   // ---------- 网络 6 ----------
   // 标题：模式传递到M区,方便使用
   // 含义：当 #SubSysMode.Mode.ManMode 为 TRUE 时置位 "ManMode_M"，否则复位（触点→线圈）
   IF #SubSysMode.Mode.ManMode THEN
       "ManMode_M" := TRUE;
   ELSE
       "ManMode_M" := FALSE;
   END_IF;
   // 含义：当 #SubSysMode.Mode.ManMode 为 TRUE 时置位 "DB1900_Communication_PC".Send.ManMode，否则复位（触点→线圈）
   IF #SubSysMode.Mode.ManMode THEN
       "DB1900_Communication_PC".Send.ManMode := TRUE;
   ELSE
       "DB1900_Communication_PC".Send.ManMode := FALSE;
   END_IF;
   // 含义：当 #SubSysMode.Mode.MastMode 为 TRUE 时置位 "MastMode_M"，否则复位（触点→线圈）
   IF #SubSysMode.Mode.MastMode THEN
       "MastMode_M" := TRUE;
   ELSE
       "MastMode_M" := FALSE;
   END_IF;
   // 含义：当 #SubSysMode.Mode.StepMode 为 TRUE 时置位 "StepMode_M"，否则复位（触点→线圈）
   IF #SubSysMode.Mode.StepMode THEN
       "StepMode_M" := TRUE;
   ELSE
       "StepMode_M" := FALSE;
   END_IF;
   // 含义：当 #SubSysMode.Mode.AutoMode 为 TRUE 时置位 "AutoMode_M"，否则复位（触点→线圈）
   IF #SubSysMode.Mode.AutoMode THEN
       "AutoMode_M" := TRUE;
   ELSE
       "AutoMode_M" := FALSE;
   END_IF;
   // 含义：当 #SubSysMode.Mode.AutoMode 为 TRUE 时置位 "DB1900_Communication_PC".Send.AutoMode，否则复位（触点→线圈）
   IF #SubSysMode.Mode.AutoMode THEN
       "DB1900_Communication_PC".Send.AutoMode := TRUE;
   ELSE
       "DB1900_Communication_PC".Send.AutoMode := FALSE;
   END_IF;
   // 含义：当 #SubSysMode.Mode.EMMode 为 TRUE 时置位 "EMMode_M"，否则复位（触点→线圈）
   IF #SubSysMode.Mode.EMMode THEN
       "EMMode_M" := TRUE;
   ELSE
       "EMMode_M" := FALSE;
   END_IF;
   // 含义：当 #SubSysMode.Mode.EMMode 为 TRUE 时置位 "DB1900_Communication_PC".Send.EmmMode，否则复位（触点→线圈）
   IF #SubSysMode.Mode.EMMode THEN
       "DB1900_Communication_PC".Send.EmmMode := TRUE;
   ELSE
       "DB1900_Communication_PC".Send.EmmMode := FALSE;
   END_IF;
   // 含义：当 #SubSysMode.Mode.StepPls 为 TRUE 时置位 "StepPls_M"，否则复位（触点→线圈）
   IF #SubSysMode.Mode.StepPls THEN
       "StepPls_M" := TRUE;
   ELSE
       "StepPls_M" := FALSE;
   END_IF;
   // 含义：当 #SubSysMode.Status.AutoModeStarted 为 TRUE 时置位 "AutoModeStarted_M"，否则复位（触点→线圈）
   IF #SubSysMode.Status.AutoModeStarted THEN
       "AutoModeStarted_M" := TRUE;
   ELSE
       "AutoModeStarted_M" := FALSE;
   END_IF;
   // 含义：当 #SubSysMode.Mode.ASMode 为 TRUE 时置位 "ASMode_M"，否则复位（触点→线圈）
   IF #SubSysMode.Mode.ASMode THEN
       "ASMode_M" := TRUE;
   ELSE
       "ASMode_M" := FALSE;
   END_IF;
   // 含义：当 #SubSysMode.Mode.ASMMode 为 TRUE 时置位 "ASMMode_M"，否则复位（触点→线圈）
   IF #SubSysMode.Mode.ASMMode THEN
       "ASMMode_M" := TRUE;
   ELSE
       "ASMMode_M" := FALSE;
   END_IF;
   // 含义：当 #SubSysMode.Mode.AllMode 为 TRUE 时置位 "AllMode_M"，否则复位（触点→线圈）
   IF #SubSysMode.Mode.AllMode THEN
       "AllMode_M" := TRUE;
   ELSE
       "AllMode_M" := FALSE;
   END_IF;
   // 含义：当 #SubSysMode.Mode.ErrRst 为 TRUE 时置位 "ErrRst_M"，否则复位（触点→线圈）
   IF #SubSysMode.Mode.ErrRst THEN
       "ErrRst_M" := TRUE;
   ELSE
       "ErrRst_M" := FALSE;
   END_IF;
   // 含义：将 #SubSysMode.Mode.ErrRst OR "DB1010_Parameter".SystemParaR.bit.ErrAutoResetOption 赋给 "ErrRst_M_Auto"
   "ErrRst_M_Auto" := #SubSysMode.Mode.ErrRst OR "DB1010_Parameter".SystemParaR.bit.ErrAutoResetOption;
   // 含义：当 "DB1010_Parameter".SystemParaR.bit.MESActive 为 TRUE 时置位 "MESConnect"，否则复位（触点→线圈）
   IF "DB1010_Parameter".SystemParaR.bit.MESActive THEN
       "MESConnect" := TRUE;
   ELSE
       "MESConnect" := FALSE;
   END_IF;

   // ---------- 网络 7 ----------
   // 标题：操作盒急停OK
   // 含义：当 NOT ("IEMOK1") 为 TRUE 时置位 "DB1148_PromptBeeper".Public.EMOK，否则复位（触点→线圈）
   IF NOT ("IEMOK1") THEN
       "DB1148_PromptBeeper".Public.EMOK := TRUE;
   ELSE
       "DB1148_PromptBeeper".Public.EMOK := FALSE;
   END_IF;
   // 含义：当 NOT ("IInsideEMOK") 为 TRUE 时置位 "DB1148_PromptBeeper".Public.InsideEMOK，否则复位（触点→线圈）
   IF NOT ("IInsideEMOK") THEN
       "DB1148_PromptBeeper".Public.InsideEMOK := TRUE;
   ELSE
       "DB1148_PromptBeeper".Public.InsideEMOK := FALSE;
   END_IF;
   // 含义：当 NOT ("IInsideEMOK1") 为 TRUE 时置位 "DB1148_PromptBeeper".Public.InsideEMOK1，否则复位（触点→线圈）
   IF NOT ("IInsideEMOK1") THEN
       "DB1148_PromptBeeper".Public.InsideEMOK1 := TRUE;
   ELSE
       "DB1148_PromptBeeper".Public.InsideEMOK1 := FALSE;
   END_IF;
   // 含义：当 NOT ("IRobotEMOK") 为 TRUE 时置位 "DB1148_PromptBeeper".Public.RobotEMOK，否则复位（触点→线圈）
   IF NOT ("IRobotEMOK") THEN
       "DB1148_PromptBeeper".Public.RobotEMOK := TRUE;
   ELSE
       "DB1148_PromptBeeper".Public.RobotEMOK := FALSE;
   END_IF;

   // ---------- 网络 8 ----------
   // 标题：调试的时候，临时关闭
   // 含义：条件 "EMMode_M" OR "DB1010_Parameter".Status.Para_ReNewEdPls OR "DB1000_StdSignal".PLS.InitialPls 成立时，将 FALSE 传送到 "Debug_True"
   IF "EMMode_M" OR "DB1010_Parameter".Status.Para_ReNewEdPls OR "DB1000_StdSignal".PLS.InitialPls THEN
       "Debug_True" := FALSE;
   END_IF;
END_FUNCTION_BLOCK

FUNCTION_BLOCK "FB1002_subSysMode"   // FB1002, SCL
{ S7_Optimized_Access := 'TRUE' }
// ============================================================
//  Block: FB1002_subSysMode
//  ============================================================
//  编号：FB1002
//  原始语言：LAD（规则翻译为 SCL）
//  含义：故障红色指示灯输出，并且存储最后的不合格状态。
   VAR_INPUT
      I_OkToStartNew : Bool;   // 可以启动新的流程
      iEMOK : Bool;   // 紧急停止OK信号
      iAirPressOK : Bool;   // 气源OK信号
      iManMode : Bool;   // 手动模式
      iAutoMode : Bool;   // 自动模式信号
      iAutoModeStart : Bool;   // 自动模式启动开关
      iBeeperQuiet : Bool;   // 蜂鸣器静音按钮
      iErrRst : Bool;   // 故障复位按钮
      iStartL : Bool;   // 左启动
      iStartR : Bool;   // 右启动
      I_ErrPresent : Bool;   // DB_ERR内有故障位存在
      I_ErrAutoReset : Bool := TRUE;   // 故障发生后自动复位。
      I_AutoRuning : Bool;   // 设备自动运行中
      I_HomeIng : Bool;   // 设备正在回原点
      I_AllStationInHomePos : Bool;   // 都在原点位置
      iHomeMode : Bool;   // 回原点按钮
      I_SP2 : Bool;   // 输入参数
   END_VAR
   VAR_OUTPUT
      oTLBlue : Bool;   // 通讯正常 塔灯-蓝
      oTLYel : Bool;   // 手动模式 塔灯-黄
      oTLGreen : Bool;   // 自动运行 塔灯-绿
      oTLRed : Bool;   // 故障报警 塔灯-红
      oTLWhite : Bool;   // 设备上电 塔灯-白
      oPanelG : Bool;   // 面板绿灯
      oPanelRed : Bool;   // 面板红灯
      oBeeper : Bool;   // 蜂鸣器
      oLightingLampClose : Bool;   // 日光灯控制
      oEMErr : Bool;   // 紧急停止故障
      oPressErr : Bool;   // 气压低故障
      oErrToBeRst : Bool;   // 发生故障，需要复位，用于屏幕提示
      oStartAutoModePrompt : Bool;   // 请启动自动模式
      oAutoModeOffPrompt : Bool;   // 自动模式已经暂停，等待循环结束！
      oEmptyMode : Bool;   // 设备进入清空模式提示信息
      oStepMode : Bool;   // 设备进入单步模式提示信息
      oModeFromTP : Bool;   // 模式来自触摸屏提示信息！
   END_VAR
   VAR
      OUT : Struct   // 静态变量
         LampTest : Bool;   // 指示灯测试
         oPanelHome : Bool;   // 面板回原点指示灯
         sp : Word;   // 静态变量
      END_STRUCT;
      Mode : Struct   // 静态变量
         ManMode : Bool;   // 手动模式
         MastMode : Bool;   // 校验模式
         StepMode : Bool;   // 单步模式
         AutoMode : Bool;   // 自动模式
         EMMode : Bool;   // 紧急停止模式
         PressLowMode : Bool;   // 气压低
         sp_1 : Bool;   // 静态变量
         sp_2 : Bool;   // 静态变量
         ASMode : Bool;   // 自动或单步模式
         ASMMode : Bool;   // 自动，单步，校验模式
         AllMode : Bool;   // 所有模式
         HomeCmd : Bool;   // 回原点命令
         ErrRst : Bool;   // 故障复位（含TPPB）
         StartPls : Bool;   // 双手启动模式使用
         StepPls : Bool;   // 双手启动模式使用
         StartLeftPls : Bool;   // 单手启动左工位
         StartRightPls : Bool;   // 单手启动右工位
         StepLeftPls : Bool;   // 单手启动左工位
         StepRightPls : Bool;   // 单手启动右工位
         ManModePls : Bool;   // 切换到手动模式脉冲
         AllModePls : Bool;   // 模式切换脉冲
         sp : DWord;   // 静态变量
      END_STRUCT;
      TPPB : Struct   // 18
         EmptyMode : Bool;   // 清空模式开始
         Bypass : Bool;   // 静态变量
         STAT6 : Bool;   // 静态变量
         STAT5 : Bool;   // 静态变量
         STAT4 : Bool;   // 静态变量
         STAT3 : Bool;   // 静态变量
         STAT2 : Bool;   // 静态变量
         STAT1 : Bool;   // 静态变量
         LampTest : Bool;   // 指示灯测试
         Home : Bool;   // 回原点
         StepMode : Bool;   // 单步按钮
         ErrRst : Bool;   // 来自触摸屏
         LampCtrol : Bool;   // ON,日光灯开
         Quiet : Bool;   // 静音，蜂鸣器
         opModeFromTP : Bool;   // 工作模式来自触摸屏选项
         sp : DWord;   // 静态变量
      END_STRUCT;
      AtTPPB : Word;   // 静态变量
      Status : Struct   // For_TP_Show
         HomePos : Bool;   // 在原点位置
         HomeIng : Bool;   // 正在原点
         AutoRunning : Bool;   // 自动运行中
         ErrPresent : Bool;   // 设备有故障
         AutoModeStarted : Bool;   // 自动模式已经启动！
      END_STRUCT;
      TPSetPageNo : Int;   // 设置当前画面号
      TPCurPageType : Int;   // 当前画面类型（工位分类）
      TPCurSubPage : Int;   // 画面子类型（手动、自动等）
      IO_FromTP : Struct   // 来自触摸屏的模拟仿真按钮输入
         spbyte : Byte;   // 来自触摸屏的模拟仿真按钮输入
         EMOK : Bool := TRUE;   // 紧急停止OK信号
         AirPressOK : Bool := TRUE;   // 气源OK信号
         ManMode : Bool;   // 手动模式
         AutoMode : Bool;   // 自动模式信号
         AutoModeStart : Bool;   // 自动模式启动开关
         ErrRst : Bool;   // 故障复位按钮
         StartLeft : Bool;   // 启动设备（左按钮）
         StartRight : Bool;   // 启动设备（右按钮）
      END_STRUCT;
      IO_Cur : Struct   // 当前实际使用的信号状态
         spbyte : Byte;   // 静态变量
         EMOK : Bool;   // 紧急停止OK信号
         AirPressOK : Bool;   // 气源OK信号
         ManMode : Bool;   // 手动模式
         AutoMode : Bool;   // 自动模式信号
         AutoModeStart : Bool;   // 自动模式启动开关
         ErrRst : Bool;   // 故障复位按钮
         StartLeft : Bool;   // 启动设备（左按钮）
         StartRight : Bool;   // 启动设备（右按钮）
      END_STRUCT;
      ModeDT : Struct   // 模式延时
         ManMode1 : Bool;   // 静态变量
         ManMode2 : Bool;   // 静态变量
         AutoMode1 : Bool;   // 静态变量
         AutoMode2 : Bool;   // 静态变量
         MastMode1 : Bool;   // 静态变量
         MastMode2 : Bool;   // 静态变量
         HomeCmd1 : Bool;   // 静态变量
         HomeCmd2 : Bool;   // 静态变量
         HomeCmd3 : Bool;   // 静态变量
         HomeCmd4 : Bool;   // 静态变量
         ErrLampOn01 : Bool;   // 静态变量
         ErrLampOn02 : Bool;   // 静态变量
      END_STRUCT;
      Aux : Struct   // 静态变量
         BeeperON_Keep : Bool;   // 静态变量
         BeeperOn : Bool;   // 静态变量
         BeeperOnPls : Bool;   // 静态变量
         ManMode : Bool;   // 用于清除触摸屏的模式选择
         ManModePls : Bool;   // 用于清除触摸屏的模式选择
         AutoMode : Bool;   // 用于清除触摸屏的模式选择
         AutoModePls : Bool;   // 用于清除触摸屏的模式选择
         ModeChangePlsHW : Bool;   // 用于记录节拍
         AutoRunningPls : Bool;   // 用于记录节拍
         OKPartPromptPls : Bool;   // 脉冲计数用
         NGPartPromptPls : Bool;   // 脉冲计数用
         ManModeOn : Bool;   // 静态变量
         AllModeOn : Bool;   // 静态变量
         AutoModeStartBtnPls : Bool;   // 静态变量
         AutoModeOnPls : Bool;   // 静态变量
         AutoModeOffCmd : Bool;   // 静态变量
         TPCurSubPage : Int;   // 静态变量
      END_STRUCT;
      Start1DT1 : IEC_TIMER;   // 静态变量
      Start1DT2 : IEC_TIMER;   // 静态变量
      Start2DT1 : IEC_TIMER;   // 静态变量
      Start2DT2 : IEC_TIMER;   // 静态变量
      xArray_SP : Array[0..91] of Byte;   // 静态变量
      lastByteAddr : Byte := 198;   // 198
      PT : Time;   // 静态变量
      ET : Time;   // 静态变量
      IN : Bool;   // 静态变量
      Q : Bool;   // 静态变量
   END_VAR
   VAR_TEMP
      T_INT : Int;   // 临时变量
   END_VAR
BEGIN

   // ---------- 网络 1 ----------
   // 标题：模拟仿真模式按钮等
   // 含义：将 (NOT (#TPPB.opModeFromTP) AND #iEMOK) OR (#TPPB.opModeFromTP AND #IO_FromTP.EMOK) 赋给 #IO_Cur.EMOK
   #IO_Cur.EMOK := (NOT (#TPPB.opModeFromTP) AND #iEMOK) OR (#TPPB.opModeFromTP AND #IO_FromTP.EMOK);
   // 含义：将 (NOT (#TPPB.opModeFromTP) AND #iAirPressOK) OR (#TPPB.opModeFromTP AND #IO_FromTP.AirPressOK) 赋给 #IO_Cur.AirPressOK
   #IO_Cur.AirPressOK := (NOT (#TPPB.opModeFromTP) AND #iAirPressOK) OR (#TPPB.opModeFromTP AND #IO_FromTP.AirPressOK);
   // 含义：将 (NOT (#TPPB.opModeFromTP) AND #iManMode) OR (#TPPB.opModeFromTP AND NOT (#IO_FromTP.AutoMode)) 赋给 #IO_Cur.ManMode
   #IO_Cur.ManMode := (NOT (#TPPB.opModeFromTP) AND #iManMode) OR (#TPPB.opModeFromTP AND NOT (#IO_FromTP.AutoMode));
   // 含义：将 (NOT (#TPPB.opModeFromTP) AND #iAutoMode) OR (#TPPB.opModeFromTP AND #IO_FromTP.AutoMode) 赋给 #IO_Cur.AutoMode
   #IO_Cur.AutoMode := (NOT (#TPPB.opModeFromTP) AND #iAutoMode) OR (#TPPB.opModeFromTP AND #IO_FromTP.AutoMode);
   // 含义：将 (NOT (#TPPB.opModeFromTP) AND #iAutoModeStart) OR (#TPPB.opModeFromTP AND #IO_FromTP.AutoModeStart) 赋给 #IO_Cur.AutoModeStart
   #IO_Cur.AutoModeStart := (NOT (#TPPB.opModeFromTP) AND #iAutoModeStart) OR (#TPPB.opModeFromTP AND #IO_FromTP.AutoModeStart);
   // 含义：将 (NOT (#TPPB.opModeFromTP) AND #iErrRst) OR (#TPPB.opModeFromTP AND #IO_FromTP.ErrRst) 赋给 #IO_Cur.ErrRst
   #IO_Cur.ErrRst := (NOT (#TPPB.opModeFromTP) AND #iErrRst) OR (#TPPB.opModeFromTP AND #IO_FromTP.ErrRst);
   // 含义：将 (NOT (#TPPB.opModeFromTP) AND #iStartL) OR (#TPPB.opModeFromTP AND #IO_FromTP.StartLeft) 赋给 #IO_Cur.StartLeft
   #IO_Cur.StartLeft := (NOT (#TPPB.opModeFromTP) AND #iStartL) OR (#TPPB.opModeFromTP AND #IO_FromTP.StartLeft);
   // 含义：将 (NOT (#TPPB.opModeFromTP) AND #iStartR) OR (#TPPB.opModeFromTP AND #IO_FromTP.StartRight) 赋给 #IO_Cur.StartRight
   #IO_Cur.StartRight := (NOT (#TPPB.opModeFromTP) AND #iStartR) OR (#TPPB.opModeFromTP AND #IO_FromTP.StartRight);
   // 含义：条件 (#iManMode OR #iAutoMode) AND NOT (#Aux.ModeChangePlsHW) 成立时，将 FALSE 传送到 #TPPB.opModeFromTP
   IF (#iManMode OR #iAutoMode) AND NOT (#Aux.ModeChangePlsHW) THEN
       #TPPB.opModeFromTP := FALSE;
   END_IF;
   // 含义：将 #iManMode OR #iAutoMode 赋给 #Aux.ModeChangePlsHW
   #Aux.ModeChangePlsHW := #iManMode OR #iAutoMode;
   // 含义：当 #TPPB.opModeFromTP 为 TRUE 时置位 #oModeFromTP，否则复位（触点→线圈）
   IF #TPPB.opModeFromTP THEN
       #oModeFromTP := TRUE;
   ELSE
       #oModeFromTP := FALSE;
   END_IF;
   // 含义：条件 #TPPB.opModeFromTP AND #iErrRst 成立时，将 FALSE 传送到 #TPPB.opModeFromTP
   IF #TPPB.opModeFromTP AND #iErrRst THEN
       #TPPB.opModeFromTP := FALSE;
   END_IF;

   // ---------- 网络 2 ----------
   // 标题：在原点位置
   // 含义：当 #I_AllStationInHomePos 为 TRUE 时置位 #Status.HomePos，否则复位（触点→线圈）
   IF #I_AllStationInHomePos THEN
       #Status.HomePos := TRUE;
   ELSE
       #Status.HomePos := FALSE;
   END_IF;
   // 含义：当 #I_HomeIng 为 TRUE 时置位 #Status.HomeIng，否则复位（触点→线圈）
   IF #I_HomeIng THEN
       #Status.HomeIng := TRUE;
   ELSE
       #Status.HomeIng := FALSE;
   END_IF;
   // 含义：当 #I_AutoRuning 为 TRUE 时置位 #Status.AutoRunning，否则复位（触点→线圈）
   IF #I_AutoRuning THEN
       #Status.AutoRunning := TRUE;
   ELSE
       #Status.AutoRunning := FALSE;
   END_IF;

   // ---------- 网络 3 ----------
   // 标题：#OUT.ErrLamp
   // 含义：当 #I_ErrPresent 为 TRUE 时置位 #Status.ErrPresent，否则复位（触点→线圈）
   IF #I_ErrPresent THEN
       #Status.ErrPresent := TRUE;
   ELSE
       #Status.ErrPresent := FALSE;
   END_IF;

   // ---------- 网络 4 ----------
   // 标题：#oTLRed
   // 注释：故障红色指示灯输出，并且存储最后的不合格状态。
   // 含义：将 #Status.ErrPresent AND #ModeDT.ErrLampOn02 赋给 #oTLRed
   #oTLRed := #Status.ErrPresent AND #ModeDT.ErrLampOn02;
   // 含义：将 ((#Status.ErrPresent AND "DB1000_StdSignal".PLS.PS05) AND #ModeDT.ErrLampOn01) OR (#Status.ErrPresent AND #ModeDT.ErrLampOn02) 赋给 #ModeDT.ErrLampOn02
   #ModeDT.ErrLampOn02 := ((#Status.ErrPresent AND "DB1000_StdSignal".PLS.PS05) AND #ModeDT.ErrLampOn01) OR (#Status.ErrPresent AND #ModeDT.ErrLampOn02);
   // 含义：将 (#Status.ErrPresent AND "DB1000_StdSignal".PLS.PS01) OR (#Status.ErrPresent AND #ModeDT.ErrLampOn01) 赋给 #ModeDT.ErrLampOn01
   #ModeDT.ErrLampOn01 := (#Status.ErrPresent AND "DB1000_StdSignal".PLS.PS01) OR (#Status.ErrPresent AND #ModeDT.ErrLampOn01);

   // ---------- 网络 5 ----------
   // 标题：#oTLYel,   #oTLGreen
   // 含义：当 #Mode.ManMode 为 TRUE 时置位 #oTLYel，否则复位（触点→线圈）
   IF #Mode.ManMode THEN
       #oTLYel := TRUE;
   ELSE
       #oTLYel := FALSE;
   END_IF;
   // 含义：将 #Mode.ASMMode AND NOT (#oTLRed) 赋给 #oTLGreen
   #oTLGreen := #Mode.ASMMode AND NOT (#oTLRed);

   // ---------- 网络 6 ----------
   // 标题：#oTLBlue
   // 含义：将 "DB720_KuKa_MainCtrl".ChangeTool.StepStart AND "DB1000_StdSignal".RectWave.Wave05 赋给 #oTLBlue
   #oTLBlue := "DB720_KuKa_MainCtrl".ChangeTool.StepStart AND "DB1000_StdSignal".RectWave.Wave05;
   // 含义：当 NOT (#Mode.EMMode) 为 TRUE 时置位 #oTLWhite，否则复位（触点→线圈）
   IF NOT (#Mode.EMMode) THEN
       #oTLWhite := TRUE;
   ELSE
       #oTLWhite := FALSE;
   END_IF;

   // ---------- 网络 7 ----------
   // 标题：#oPanelG
   // 含义：将 ((((#Status.HomeIng AND "DB1000_StdSignal".RectWave.Wave02) AND NOT (TRUE)) OR (((((#Mode.AutoMode AND NOT (#I_HomeIng)) AND NOT (#Status.AutoRunning)) AND NOT (#Status.AutoModeStarted)) AND #Status.HomePos) AND "DB1000_StdSignal".RectWave.Wave05) OR #Status.AutoModeStarted OR ("AutoMode_M" AND "DB1900_Communication_PC".Send.DrillRunning)) AND NOT (#Aux.AutoModeOffCmd)) OR (#Aux.AutoModeOffCmd AND "DB1000_StdSignal".PLS.PS02) 赋给 #oPanelG
   #oPanelG := ((((#Status.HomeIng AND "DB1000_StdSignal".RectWave.Wave02) AND NOT (TRUE)) OR (((((#Mode.AutoMode AND NOT (#I_HomeIng)) AND NOT (#Status.AutoRunning)) AND NOT (#Status.AutoModeStarted)) AND #Status.HomePos) AND "DB1000_StdSignal".RectWave.Wave05) OR #Status.AutoModeStarted OR ("AutoMode_M" AND "DB1900_Communication_PC".Send.DrillRunning)) AND NOT (#Aux.AutoModeOffCmd)) OR (#Aux.AutoModeOffCmd AND "DB1000_StdSignal".PLS.PS02);

   // ---------- 网络 8 ----------
   // 标题：#oPanelRed
   // 注释：故障红色指示灯输出，并且存储最后的不合格状态。
   // 含义：将 #oTLRed OR (#I_HomeIng AND "DB1000_StdSignal".RectWave.Wave02) 赋给 #oPanelRed
   #oPanelRed := #oTLRed OR (#I_HomeIng AND "DB1000_StdSignal".RectWave.Wave02);

   // ---------- 网络 9 ----------
   // 标题：#oBeeper
   // 含义：将 #oTLRed AND NOT (#Aux.BeeperOn) 赋给 #Aux.BeeperOnPls
   #Aux.BeeperOnPls := #oTLRed AND NOT (#Aux.BeeperOn);
   // 含义：当 #oTLRed 为 TRUE 时置位 #Aux.BeeperOn，否则复位（触点→线圈）
   IF #oTLRed THEN
       #Aux.BeeperOn := TRUE;
   ELSE
       #Aux.BeeperOn := FALSE;
   END_IF;
   // 含义：将 (((#oTLRed AND #Aux.BeeperOnPls) OR (#oTLRed AND #Aux.BeeperON_Keep)) AND NOT (#Mode.ErrRst)) AND NOT (#iBeeperQuiet) 赋给 #Aux.BeeperON_Keep
   #Aux.BeeperON_Keep := (((#oTLRed AND #Aux.BeeperOnPls) OR (#oTLRed AND #Aux.BeeperON_Keep)) AND NOT (#Mode.ErrRst)) AND NOT (#iBeeperQuiet);
   // 含义：将 (((#oTLRed AND #Aux.BeeperOnPls) OR (#oTLRed AND #Aux.BeeperON_Keep)) AND "DB1000_StdSignal".RectWave.Beeper) AND NOT (#TPPB.Quiet) 赋给 #oBeeper
   #oBeeper := (((#oTLRed AND #Aux.BeeperOnPls) OR (#oTLRed AND #Aux.BeeperON_Keep)) AND "DB1000_StdSignal".RectWave.Beeper) AND NOT (#TPPB.Quiet);

   // ---------- 网络 10 ----------
   // 标题：#oPanelHome
   // 含义：将 (#Status.HomeIng AND "DB1000_StdSignal".RectWave.Wave02) OR #I_AllStationInHomePos 赋给 #OUT.oPanelHome
   #OUT.oPanelHome := (#Status.HomeIng AND "DB1000_StdSignal".RectWave.Wave02) OR #I_AllStationInHomePos;

   // ---------- 网络 11 ----------
   // 标题：#oErrToBeRst
   // 含义：将 (((#oTLRed OR #oErrToBeRst) AND NOT (#Mode.ErrRst)) AND NOT (#I_ErrAutoReset)) AND #Mode.AllMode 赋给 #oErrToBeRst
   #oErrToBeRst := (((#oTLRed OR #oErrToBeRst) AND NOT (#Mode.ErrRst)) AND NOT (#I_ErrAutoReset)) AND #Mode.AllMode;

   // ---------- 网络 12 ----------
   // 标题：#oEMErr,   #oPressErr
   // 含义：当 NOT (#IO_Cur.EMOK) 为 TRUE 时置位 #oEMErr，否则复位（触点→线圈）
   IF NOT (#IO_Cur.EMOK) THEN
       #oEMErr := TRUE;
   ELSE
       #oEMErr := FALSE;
   END_IF;
   // 含义：条件 #IO_Cur.EMOK AND NOT (#IO_Cur.AirPressOK) 成立时，将 TRUE 传送到 #oPressErr
   IF #IO_Cur.EMOK AND NOT (#IO_Cur.AirPressOK) THEN
       #oPressErr := TRUE;
   END_IF;
   // 含义：条件 #Mode.ErrRst AND #IO_Cur.AirPressOK 成立时，将 FALSE 传送到 #oPressErr
   IF #Mode.ErrRst AND #IO_Cur.AirPressOK THEN
       #oPressErr := FALSE;
   END_IF;

   // ---------- 网络 13 ----------
   // 标题：Mode ChangePls;
   // 含义：将 #IO_Cur.ManMode AND NOT (#Aux.ManMode) 赋给 #Aux.ManModePls
   #Aux.ManModePls := #IO_Cur.ManMode AND NOT (#Aux.ManMode);
   // 含义：当 #IO_Cur.ManMode 为 TRUE 时置位 #Aux.ManMode，否则复位（触点→线圈）
   IF #IO_Cur.ManMode THEN
       #Aux.ManMode := TRUE;
   ELSE
       #Aux.ManMode := FALSE;
   END_IF;
   // 含义：将 #IO_Cur.AutoMode AND NOT (#Aux.AutoMode) 赋给 #Aux.AutoModePls
   #Aux.AutoModePls := #IO_Cur.AutoMode AND NOT (#Aux.AutoMode);
   // 含义：当 #IO_Cur.AutoMode 为 TRUE 时置位 #Aux.AutoMode，否则复位（触点→线圈）
   IF #IO_Cur.AutoMode THEN
       #Aux.AutoMode := TRUE;
   ELSE
       #Aux.AutoMode := FALSE;
   END_IF;

   // ---------- 网络 14 ----------
   // 标题：模式延时处理。
   // 含义：将 (((((("DB1000_StdSignal".PowerOn AND NOT (#oEMErr)) AND NOT (#oPressErr)) AND #IO_Cur.ManMode) AND NOT (#IO_Cur.AutoMode)) AND "DB1000_StdSignal".PLS.PS01) AND #ModeDT.ManMode1) OR ((((("DB1000_StdSignal".PowerOn AND NOT (#oEMErr)) AND NOT (#oPressErr)) AND #IO_Cur.ManMode) AND NOT (#IO_Cur.AutoMode)) AND #ModeDT.ManMode2) 赋给 #ModeDT.ManMode2
   #ModeDT.ManMode2 := (((((("DB1000_StdSignal".PowerOn AND NOT (#oEMErr)) AND NOT (#oPressErr)) AND #IO_Cur.ManMode) AND NOT (#IO_Cur.AutoMode)) AND "DB1000_StdSignal".PLS.PS01) AND #ModeDT.ManMode1) OR ((((("DB1000_StdSignal".PowerOn AND NOT (#oEMErr)) AND NOT (#oPressErr)) AND #IO_Cur.ManMode) AND NOT (#IO_Cur.AutoMode)) AND #ModeDT.ManMode2);
   // 含义：将 ((((("DB1000_StdSignal".PowerOn AND NOT (#oEMErr)) AND NOT (#oPressErr)) AND #IO_Cur.ManMode) AND NOT (#IO_Cur.AutoMode)) AND "DB1000_StdSignal".PLS.PS01) OR ((((("DB1000_StdSignal".PowerOn AND NOT (#oEMErr)) AND NOT (#oPressErr)) AND #IO_Cur.ManMode) AND NOT (#IO_Cur.AutoMode)) AND #ModeDT.ManMode1) 赋给 #ModeDT.ManMode1
   #ModeDT.ManMode1 := ((((("DB1000_StdSignal".PowerOn AND NOT (#oEMErr)) AND NOT (#oPressErr)) AND #IO_Cur.ManMode) AND NOT (#IO_Cur.AutoMode)) AND "DB1000_StdSignal".PLS.PS01) OR ((((("DB1000_StdSignal".PowerOn AND NOT (#oEMErr)) AND NOT (#oPressErr)) AND #IO_Cur.ManMode) AND NOT (#IO_Cur.AutoMode)) AND #ModeDT.ManMode1);
   // 含义：将 (((((("DB1000_StdSignal".PowerOn AND NOT (#oEMErr)) AND NOT (#oPressErr)) AND NOT (#IO_Cur.ManMode)) AND #IO_Cur.AutoMode) AND "DB1000_StdSignal".PLS.PS01) AND #ModeDT.AutoMode1) OR ((((("DB1000_StdSignal".PowerOn AND NOT (#oEMErr)) AND NOT (#oPressErr)) AND NOT (#IO_Cur.ManMode)) AND #IO_Cur.AutoMode) AND #ModeDT.AutoMode2) 赋给 #ModeDT.AutoMode2
   #ModeDT.AutoMode2 := (((((("DB1000_StdSignal".PowerOn AND NOT (#oEMErr)) AND NOT (#oPressErr)) AND NOT (#IO_Cur.ManMode)) AND #IO_Cur.AutoMode) AND "DB1000_StdSignal".PLS.PS01) AND #ModeDT.AutoMode1) OR ((((("DB1000_StdSignal".PowerOn AND NOT (#oEMErr)) AND NOT (#oPressErr)) AND NOT (#IO_Cur.ManMode)) AND #IO_Cur.AutoMode) AND #ModeDT.AutoMode2);
   // 含义：将 ((((("DB1000_StdSignal".PowerOn AND NOT (#oEMErr)) AND NOT (#oPressErr)) AND NOT (#IO_Cur.ManMode)) AND #IO_Cur.AutoMode) AND "DB1000_StdSignal".PLS.PS01) OR ((((("DB1000_StdSignal".PowerOn AND NOT (#oEMErr)) AND NOT (#oPressErr)) AND NOT (#IO_Cur.ManMode)) AND #IO_Cur.AutoMode) AND #ModeDT.AutoMode1) 赋给 #ModeDT.AutoMode1
   #ModeDT.AutoMode1 := ((((("DB1000_StdSignal".PowerOn AND NOT (#oEMErr)) AND NOT (#oPressErr)) AND NOT (#IO_Cur.ManMode)) AND #IO_Cur.AutoMode) AND "DB1000_StdSignal".PLS.PS01) OR ((((("DB1000_StdSignal".PowerOn AND NOT (#oEMErr)) AND NOT (#oPressErr)) AND NOT (#IO_Cur.ManMode)) AND #IO_Cur.AutoMode) AND #ModeDT.AutoMode1);
   // 含义：将 (((((("DB1000_StdSignal".PowerOn AND NOT (#oEMErr)) AND NOT (#oPressErr)) AND NOT (#IO_Cur.ManMode)) AND NOT (#IO_Cur.AutoMode)) AND "DB1000_StdSignal".PLS.PS01) AND #ModeDT.MastMode1) OR ((((("DB1000_StdSignal".PowerOn AND NOT (#oEMErr)) AND NOT (#oPressErr)) AND NOT (#IO_Cur.ManMode)) AND NOT (#IO_Cur.AutoMode)) AND #ModeDT.MastMode2) 赋给 #ModeDT.MastMode2
   #ModeDT.MastMode2 := (((((("DB1000_StdSignal".PowerOn AND NOT (#oEMErr)) AND NOT (#oPressErr)) AND NOT (#IO_Cur.ManMode)) AND NOT (#IO_Cur.AutoMode)) AND "DB1000_StdSignal".PLS.PS01) AND #ModeDT.MastMode1) OR ((((("DB1000_StdSignal".PowerOn AND NOT (#oEMErr)) AND NOT (#oPressErr)) AND NOT (#IO_Cur.ManMode)) AND NOT (#IO_Cur.AutoMode)) AND #ModeDT.MastMode2);
   // 含义：将 ((((("DB1000_StdSignal".PowerOn AND NOT (#oEMErr)) AND NOT (#oPressErr)) AND NOT (#IO_Cur.ManMode)) AND NOT (#IO_Cur.AutoMode)) AND "DB1000_StdSignal".PLS.PS01) OR ((((("DB1000_StdSignal".PowerOn AND NOT (#oEMErr)) AND NOT (#oPressErr)) AND NOT (#IO_Cur.ManMode)) AND NOT (#IO_Cur.AutoMode)) AND #ModeDT.MastMode1) 赋给 #ModeDT.MastMode1
   #ModeDT.MastMode1 := ((((("DB1000_StdSignal".PowerOn AND NOT (#oEMErr)) AND NOT (#oPressErr)) AND NOT (#IO_Cur.ManMode)) AND NOT (#IO_Cur.AutoMode)) AND "DB1000_StdSignal".PLS.PS01) OR ((((("DB1000_StdSignal".PowerOn AND NOT (#oEMErr)) AND NOT (#oPressErr)) AND NOT (#IO_Cur.ManMode)) AND NOT (#IO_Cur.AutoMode)) AND #ModeDT.MastMode1);
   // 含义：将 (((((("DB1000_StdSignal".PowerOn AND NOT (#oEMErr)) AND NOT (#oPressErr)) AND #Mode.ErrRst) OR ((("DB1000_StdSignal".PowerOn AND NOT (#oEMErr)) AND NOT (#oPressErr)) AND #iHomeMode)) AND "DB1000_StdSignal".PLS.PS05) AND #ModeDT.HomeCmd3) OR ((((("DB1000_StdSignal".PowerOn AND NOT (#oEMErr)) AND NOT (#oPressErr)) AND #Mode.ErrRst) OR ((("DB1000_StdSignal".PowerOn AND NOT (#oEMErr)) AND NOT (#oPressErr)) AND #iHomeMode)) AND #ModeDT.HomeCmd4) 赋给 #ModeDT.HomeCmd4
   #ModeDT.HomeCmd4 := (((((("DB1000_StdSignal".PowerOn AND NOT (#oEMErr)) AND NOT (#oPressErr)) AND #Mode.ErrRst) OR ((("DB1000_StdSignal".PowerOn AND NOT (#oEMErr)) AND NOT (#oPressErr)) AND #iHomeMode)) AND "DB1000_StdSignal".PLS.PS05) AND #ModeDT.HomeCmd3) OR ((((("DB1000_StdSignal".PowerOn AND NOT (#oEMErr)) AND NOT (#oPressErr)) AND #Mode.ErrRst) OR ((("DB1000_StdSignal".PowerOn AND NOT (#oEMErr)) AND NOT (#oPressErr)) AND #iHomeMode)) AND #ModeDT.HomeCmd4);
   // 含义：将 (((((("DB1000_StdSignal".PowerOn AND NOT (#oEMErr)) AND NOT (#oPressErr)) AND #Mode.ErrRst) OR ((("DB1000_StdSignal".PowerOn AND NOT (#oEMErr)) AND NOT (#oPressErr)) AND #iHomeMode)) AND "DB1000_StdSignal".PLS.PS05) AND #ModeDT.HomeCmd2) OR ((((("DB1000_StdSignal".PowerOn AND NOT (#oEMErr)) AND NOT (#oPressErr)) AND #Mode.ErrRst) OR ((("DB1000_StdSignal".PowerOn AND NOT (#oEMErr)) AND NOT (#oPressErr)) AND #iHomeMode)) AND #ModeDT.HomeCmd3) 赋给 #ModeDT.HomeCmd3
   #ModeDT.HomeCmd3 := (((((("DB1000_StdSignal".PowerOn AND NOT (#oEMErr)) AND NOT (#oPressErr)) AND #Mode.ErrRst) OR ((("DB1000_StdSignal".PowerOn AND NOT (#oEMErr)) AND NOT (#oPressErr)) AND #iHomeMode)) AND "DB1000_StdSignal".PLS.PS05) AND #ModeDT.HomeCmd2) OR ((((("DB1000_StdSignal".PowerOn AND NOT (#oEMErr)) AND NOT (#oPressErr)) AND #Mode.ErrRst) OR ((("DB1000_StdSignal".PowerOn AND NOT (#oEMErr)) AND NOT (#oPressErr)) AND #iHomeMode)) AND #ModeDT.HomeCmd3);
   // 含义：将 (((((("DB1000_StdSignal".PowerOn AND NOT (#oEMErr)) AND NOT (#oPressErr)) AND #Mode.ErrRst) OR ((("DB1000_StdSignal".PowerOn AND NOT (#oEMErr)) AND NOT (#oPressErr)) AND #iHomeMode)) AND "DB1000_StdSignal".PLS.PS10) AND #ModeDT.HomeCmd1) OR ((((("DB1000_StdSignal".PowerOn AND NOT (#oEMErr)) AND NOT (#oPressErr)) AND #Mode.ErrRst) OR ((("DB1000_StdSignal".PowerOn AND NOT (#oEMErr)) AND NOT (#oPressErr)) AND #iHomeMode)) AND #ModeDT.HomeCmd2) 赋给 #ModeDT.HomeCmd2
   #ModeDT.HomeCmd2 := (((((("DB1000_StdSignal".PowerOn AND NOT (#oEMErr)) AND NOT (#oPressErr)) AND #Mode.ErrRst) OR ((("DB1000_StdSignal".PowerOn AND NOT (#oEMErr)) AND NOT (#oPressErr)) AND #iHomeMode)) AND "DB1000_StdSignal".PLS.PS10) AND #ModeDT.HomeCmd1) OR ((((("DB1000_StdSignal".PowerOn AND NOT (#oEMErr)) AND NOT (#oPressErr)) AND #Mode.ErrRst) OR ((("DB1000_StdSignal".PowerOn AND NOT (#oEMErr)) AND NOT (#oPressErr)) AND #iHomeMode)) AND #ModeDT.HomeCmd2);
   // 含义：将 ((((("DB1000_StdSignal".PowerOn AND NOT (#oEMErr)) AND NOT (#oPressErr)) AND #Mode.ErrRst) OR ((("DB1000_StdSignal".PowerOn AND NOT (#oEMErr)) AND NOT (#oPressErr)) AND #iHomeMode)) AND "DB1000_StdSignal".PLS.PS10) OR ((((("DB1000_StdSignal".PowerOn AND NOT (#oEMErr)) AND NOT (#oPressErr)) AND #Mode.ErrRst) OR ((("DB1000_StdSignal".PowerOn AND NOT (#oEMErr)) AND NOT (#oPressErr)) AND #iHomeMode)) AND #ModeDT.HomeCmd1) 赋给 #ModeDT.HomeCmd1
   #ModeDT.HomeCmd1 := ((((("DB1000_StdSignal".PowerOn AND NOT (#oEMErr)) AND NOT (#oPressErr)) AND #Mode.ErrRst) OR ((("DB1000_StdSignal".PowerOn AND NOT (#oEMErr)) AND NOT (#oPressErr)) AND #iHomeMode)) AND "DB1000_StdSignal".PLS.PS10) OR ((((("DB1000_StdSignal".PowerOn AND NOT (#oEMErr)) AND NOT (#oPressErr)) AND #Mode.ErrRst) OR ((("DB1000_StdSignal".PowerOn AND NOT (#oEMErr)) AND NOT (#oPressErr)) AND #iHomeMode)) AND #ModeDT.HomeCmd1);

   // ---------- 网络 15 ----------
   // 标题：AutoMode Push On
   // 含义：将 (((#Mode.ASMode AND #IO_Cur.AutoModeStart) AND NOT (#Aux.AutoModeStartBtnPls)) AND NOT (#Status.AutoModeStarted)) OR (((#Mode.ASMode AND #IO_Cur.AutoModeStart) AND NOT (#Aux.AutoModeStartBtnPls)) AND #Aux.AutoModeOffCmd) 赋给 #Aux.AutoModeOnPls
   #Aux.AutoModeOnPls := (((#Mode.ASMode AND #IO_Cur.AutoModeStart) AND NOT (#Aux.AutoModeStartBtnPls)) AND NOT (#Status.AutoModeStarted)) OR (((#Mode.ASMode AND #IO_Cur.AutoModeStart) AND NOT (#Aux.AutoModeStartBtnPls)) AND #Aux.AutoModeOffCmd);
   // 含义：条件 (((#Mode.ASMode AND #IO_Cur.AutoModeStart) AND NOT (#Aux.AutoModeStartBtnPls)) AND NOT (#Status.AutoModeStarted)) OR (((#Mode.ASMode AND #IO_Cur.AutoModeStart) AND NOT (#Aux.AutoModeStartBtnPls)) AND #Aux.AutoModeOffCmd) 成立时，将 FALSE 传送到 #Aux.AutoModeOffCmd
   IF (((#Mode.ASMode AND #IO_Cur.AutoModeStart) AND NOT (#Aux.AutoModeStartBtnPls)) AND NOT (#Status.AutoModeStarted)) OR (((#Mode.ASMode AND #IO_Cur.AutoModeStart) AND NOT (#Aux.AutoModeStartBtnPls)) AND #Aux.AutoModeOffCmd) THEN
       #Aux.AutoModeOffCmd := FALSE;
   END_IF;
   // 含义：条件 (((#Mode.ASMode AND #IO_Cur.AutoModeStart) AND NOT (#Aux.AutoModeStartBtnPls)) AND NOT (#Status.AutoModeStarted)) OR (((#Mode.ASMode AND #IO_Cur.AutoModeStart) AND NOT (#Aux.AutoModeStartBtnPls)) AND #Aux.AutoModeOffCmd) 成立时，将 FALSE 传送到 #TPPB.StepMode
   IF (((#Mode.ASMode AND #IO_Cur.AutoModeStart) AND NOT (#Aux.AutoModeStartBtnPls)) AND NOT (#Status.AutoModeStarted)) OR (((#Mode.ASMode AND #IO_Cur.AutoModeStart) AND NOT (#Aux.AutoModeStartBtnPls)) AND #Aux.AutoModeOffCmd) THEN
       #TPPB.StepMode := FALSE;
   END_IF;
   // 含义：条件 (((#Mode.ASMode AND #IO_Cur.AutoModeStart) AND NOT (#Aux.AutoModeStartBtnPls)) AND NOT (#Aux.AutoModeOnPls)) AND #Status.AutoModeStarted 成立时，将 TRUE 传送到 #Aux.AutoModeOffCmd
   IF (((#Mode.ASMode AND #IO_Cur.AutoModeStart) AND NOT (#Aux.AutoModeStartBtnPls)) AND NOT (#Aux.AutoModeOnPls)) AND #Status.AutoModeStarted THEN
       #Aux.AutoModeOffCmd := TRUE;
   END_IF;
   // 含义：将 #Mode.ASMode AND #IO_Cur.AutoModeStart 赋给 #Aux.AutoModeStartBtnPls
   #Aux.AutoModeStartBtnPls := #Mode.ASMode AND #IO_Cur.AutoModeStart;
   // 含义：将 #Mode.ASMode AND #Aux.AutoModeOffCmd 赋给 #oAutoModeOffPrompt
   #oAutoModeOffPrompt := #Mode.ASMode AND #Aux.AutoModeOffCmd;
   // 含义：条件 NOT (#Status.AutoModeStarted) AND NOT (#Status.AutoRunning) 成立时，将 FALSE 传送到 #Aux.AutoModeOffCmd
   IF NOT (#Status.AutoModeStarted) AND NOT (#Status.AutoRunning) THEN
       #Aux.AutoModeOffCmd := FALSE;
   END_IF;

   // ---------- 网络 16 ----------
   // 标题：自动模式已经启动！
   // 含义：将 (((((((#Mode.AutoMode AND #Aux.AutoModeOnPls) AND #Status.HomePos) AND #I_OkToStartNew) AND NOT (#I_AutoRuning)) AND NOT (#I_HomeIng)) OR (#Mode.AutoMode AND #Status.AutoModeStarted)) AND NOT (#TPPB.StepMode)) AND NOT (#Aux.AutoModeOffCmd) 赋给 #Status.AutoModeStarted
   #Status.AutoModeStarted := (((((((#Mode.AutoMode AND #Aux.AutoModeOnPls) AND #Status.HomePos) AND #I_OkToStartNew) AND NOT (#I_AutoRuning)) AND NOT (#I_HomeIng)) OR (#Mode.AutoMode AND #Status.AutoModeStarted)) AND NOT (#TPPB.StepMode)) AND NOT (#Aux.AutoModeOffCmd);
   // 含义：将 (#Mode.AutoMode AND NOT (#Status.AutoModeStarted)) AND NOT (#Status.AutoRunning) 赋给 #oStartAutoModePrompt
   #oStartAutoModePrompt := (#Mode.AutoMode AND NOT (#Status.AutoModeStarted)) AND NOT (#Status.AutoRunning);

   // ---------- 网络 17 ----------
   // 标题：5种模式，用于触摸屏显示
   // 含义：当 #ModeDT.ManMode2 为 TRUE 时置位 #Mode.ManMode，否则复位（触点→线圈）
   IF #ModeDT.ManMode2 THEN
       #Mode.ManMode := TRUE;
   ELSE
       #Mode.ManMode := FALSE;
   END_IF;
   // 含义：将 #ModeDT.AutoMode2 AND NOT (#TPPB.StepMode) 赋给 #Mode.AutoMode
   #Mode.AutoMode := #ModeDT.AutoMode2 AND NOT (#TPPB.StepMode);
   // 含义：将 #ModeDT.AutoMode2 AND #TPPB.StepMode 赋给 #Mode.StepMode
   #Mode.StepMode := #ModeDT.AutoMode2 AND #TPPB.StepMode;
   // 含义：当 #ModeDT.MastMode2 为 TRUE 时置位 #Mode.MastMode，否则复位（触点→线圈）
   IF #ModeDT.MastMode2 THEN
       #Mode.MastMode := TRUE;
   ELSE
       #Mode.MastMode := FALSE;
   END_IF;
   // 含义：当 #oEMErr 为 TRUE 时置位 #Mode.EMMode，否则复位（触点→线圈）
   IF #oEMErr THEN
       #Mode.EMMode := TRUE;
   ELSE
       #Mode.EMMode := FALSE;
   END_IF;
   // 含义：将 NOT (#Mode.EMMode) AND #oPressErr 赋给 #Mode.PressLowMode
   #Mode.PressLowMode := NOT (#Mode.EMMode) AND #oPressErr;

   // ---------- 网络 18 ----------
   // 标题：模式整合，用于程序中，与触摸屏无关
   // 含义：将 #Mode.AutoMode OR #Mode.StepMode 赋给 #Mode.ASMode
   #Mode.ASMode := #Mode.AutoMode OR #Mode.StepMode;
   // 含义：将 #Mode.ASMode OR #Mode.MastMode 赋给 #Mode.ASMMode
   #Mode.ASMMode := #Mode.ASMode OR #Mode.MastMode;
   // 含义：将 #Mode.ManMode OR #Mode.ASMMode 赋给 #Mode.AllMode
   #Mode.AllMode := #Mode.ManMode OR #Mode.ASMMode;
   // 含义：将 #ModeDT.HomeCmd2 OR #TPPB.Home 赋给 #Mode.HomeCmd
   #Mode.HomeCmd := #ModeDT.HomeCmd2 OR #TPPB.Home;
   // 含义：将 #IO_Cur.ErrRst OR #TPPB.ErrRst 赋给 #Mode.ErrRst
   #Mode.ErrRst := #IO_Cur.ErrRst OR #TPPB.ErrRst;

   // ---------- 网络 19 ----------
   // 标题：切换到手动模式脉冲
   // 含义：将 #Mode.ManMode AND NOT (#Aux.ManModeOn) 赋给 #Mode.ManModePls
   #Mode.ManModePls := #Mode.ManMode AND NOT (#Aux.ManModeOn);
   // 含义：当 #Mode.ManMode 为 TRUE 时置位 #Aux.ManModeOn，否则复位（触点→线圈）
   IF #Mode.ManMode THEN
       #Aux.ManModeOn := TRUE;
   ELSE
       #Aux.ManModeOn := FALSE;
   END_IF;
   // 含义：将 #Mode.AllMode AND NOT (#Aux.AllModeOn) 赋给 #Mode.AllModePls
   #Mode.AllModePls := #Mode.AllMode AND NOT (#Aux.AllModeOn);
   // 含义：当 #Mode.AllMode 为 TRUE 时置位 #Aux.AllModeOn，否则复位（触点→线圈）
   IF #Mode.AllMode THEN
       #Aux.AllModeOn := TRUE;
   ELSE
       #Aux.AllModeOn := FALSE;
   END_IF;

   // ---------- 网络 20 ----------
   // 标题：TPPB 清除；
   // 含义：条件 NOT (#Mode.AllMode) 成立时，将 FALSE 传送到 #TPPB.Home
   IF NOT (#Mode.AllMode) THEN
       #TPPB.Home := FALSE;
   END_IF;
   // 含义：条件 NOT (#Mode.AllMode) 成立时，将 FALSE 传送到 #TPPB.ErrRst
   IF NOT (#Mode.AllMode) THEN
       #TPPB.ErrRst := FALSE;
   END_IF;
   // 含义：条件 NOT (#Mode.AllMode) 成立时，将 FALSE 传送到 #TPPB.StepMode
   IF NOT (#Mode.AllMode) THEN
       #TPPB.StepMode := FALSE;
   END_IF;

   // ---------- 网络 21 ----------
   // 标题：启动延时
   // 注释：启动信号，考虑双工位情况，如果单工位，可以只用其中之一的启动，如果是双手启动
   // ，则都用上，万能！！！
   // 含义：调用计数器实例 #Start1DT1.TON（上升沿计数，当前值写入 CV）
   #Start1DT1.TON(IN := #IO_Cur.StartLeft,
                  PT := t#30ms);
   // 含义：调用计数器实例 #Start1DT2.TON（上升沿计数，当前值写入 CV）
   #Start1DT2.TON(IN := #IO_Cur.StartLeft,
                  PT := t#130ms);
   // 含义：调用计数器实例 #Start2DT1.TON（上升沿计数，当前值写入 CV）
   #Start2DT1.TON(IN := #IO_Cur.StartRight,
                  PT := t#30ms);
   // 含义：调用计数器实例 #Start2DT2.TON（上升沿计数，当前值写入 CV）
   #Start2DT2.TON(IN := #IO_Cur.StartRight,
                  PT := t#130ms);
   // 含义：将 #Start1DT1.Q AND NOT (#Start1DT2.Q) 赋给 #Mode.StartLeftPls
   #Mode.StartLeftPls := #Start1DT1.Q AND NOT (#Start1DT2.Q);
   // 含义：将 #Start2DT1.Q AND NOT (#Start2DT2.Q) 赋给 #Mode.StartRightPls
   #Mode.StartRightPls := #Start2DT1.Q AND NOT (#Start2DT2.Q);
   // 含义：将 #Mode.StartLeftPls AND #Mode.StartRightPls 赋给 #Mode.StartPls
   #Mode.StartPls := #Mode.StartLeftPls AND #Mode.StartRightPls;

   // ---------- 网络 22 ----------
   // 标题：单步脉冲
   // 注释：单步信号，考虑双工位情况，如果单工位，可以只用其中之一的启动，如果是双手启动
   // ，则都用上，万能！！！   发生故障后，需要复位自动才会继续
   // 含义：将 (NOT (#oErrToBeRst) AND NOT (#Mode.StepMode)) OR (NOT (#oErrToBeRst) AND #Mode.StartLeftPls) 赋给 #Mode.StepLeftPls
   #Mode.StepLeftPls := (NOT (#oErrToBeRst) AND NOT (#Mode.StepMode)) OR (NOT (#oErrToBeRst) AND #Mode.StartLeftPls);
   // 含义：将 (NOT (#oErrToBeRst) AND NOT (#Mode.StepMode)) OR (NOT (#oErrToBeRst) AND #Mode.StartRightPls) 赋给 #Mode.StepRightPls
   #Mode.StepRightPls := (NOT (#oErrToBeRst) AND NOT (#Mode.StepMode)) OR (NOT (#oErrToBeRst) AND #Mode.StartRightPls);
   // 含义：将 ((NOT (#oErrToBeRst) AND #Mode.StepLeftPls) OR (NOT (#oErrToBeRst) AND #Mode.StepRightPls)) AND NOT (#oErrToBeRst) 赋给 #Mode.StepPls
   #Mode.StepPls := ((NOT (#oErrToBeRst) AND #Mode.StepLeftPls) OR (NOT (#oErrToBeRst) AND #Mode.StepRightPls)) AND NOT (#oErrToBeRst);

   // ---------- 网络 23 ----------
   // 标题：模式切换时页面切换；
   // 含义：条件 (((NOT (#TPPB.opModeFromTP) AND #IO_Cur.EMOK) AND #IO_Cur.AirPressOK) AND #IO_Cur.ManMode) AND NOT (#Mode.ManMode) 成立时，将 100 传送到 #TPSetPageNo
   IF (((NOT (#TPPB.opModeFromTP) AND #IO_Cur.EMOK) AND #IO_Cur.AirPressOK) AND #IO_Cur.ManMode) AND NOT (#Mode.ManMode) THEN
       #TPSetPageNo := 100;
   END_IF;
   // 含义：条件 (((NOT (#TPPB.opModeFromTP) AND #IO_Cur.EMOK) AND #IO_Cur.AirPressOK) AND #IO_Cur.AutoMode) AND NOT (#Mode.ASMMode) 成立时，将 200 传送到 #TPSetPageNo
   IF (((NOT (#TPPB.opModeFromTP) AND #IO_Cur.EMOK) AND #IO_Cur.AirPressOK) AND #IO_Cur.AutoMode) AND NOT (#Mode.ASMMode) THEN
       #TPSetPageNo := 200;
   END_IF;
   // 含义：条件 ((NOT (#TPPB.opModeFromTP) AND #IO_Cur.EMOK) AND #IO_Cur.AirPressOK) AND #Mode.MastMode 成立时，将 240 传送到 #TPSetPageNo
   IF ((NOT (#TPPB.opModeFromTP) AND #IO_Cur.EMOK) AND #IO_Cur.AirPressOK) AND #Mode.MastMode THEN
       #TPSetPageNo := 240;
   END_IF;
   // 含义：条件 "DB1000_StdSignal".PLS.InitialPls 成立时，将 1 传送到 #TPSetPageNo
   IF "DB1000_StdSignal".PLS.InitialPls THEN
       #TPSetPageNo := 1;
   END_IF;
   // 含义：条件 (#TPCurSubPage <> #Aux.TPCurSubPage) 成立时，将 #TPCurSubPage 传送到 #Aux.TPCurSubPage
   IF (#TPCurSubPage <> #Aux.TPCurSubPage) THEN
       #Aux.TPCurSubPage := #TPCurSubPage;
   END_IF;
   // 含义：条件 (#TPCurSubPage <> #Aux.TPCurSubPage) 成立时，将 (#TPCurSubPage + #TPCurPageType) 传送到 #TPSetPageNo
   IF (#TPCurSubPage <> #Aux.TPCurSubPage) THEN
       #TPSetPageNo := (#TPCurSubPage + #TPCurPageType);
   END_IF;
   // 含义：将 (#TPSetPageNo / 100) 赋给 #T_INT
   #T_INT := (#TPSetPageNo / 100);
   // 含义：将 (#T_INT * 100) 赋给 #TPCurPageType
   #TPCurPageType := (#T_INT * 100);
   // 含义：将 (#TPSetPageNo - #TPCurPageType) 赋给 #TPCurSubPage
   #TPCurSubPage := (#TPSetPageNo - #TPCurPageType);

   // ---------- 网络 24 ----------
   // 标题：#OUT.LampTest
   // 含义：将 #TPPB.LampTest OR "DB1000_StdSignal".LampTest 赋给 #OUT.LampTest
   #OUT.LampTest := #TPPB.LampTest OR "DB1000_StdSignal".LampTest;
   // 含义：条件 #TPPB.LampTest OR "DB1000_StdSignal".LampTest 成立时，将 TRUE 传送到 #oTLRed
   IF #TPPB.LampTest OR "DB1000_StdSignal".LampTest THEN
       #oTLRed := TRUE;
   END_IF;
   // 含义：条件 #TPPB.LampTest OR "DB1000_StdSignal".LampTest 成立时，将 TRUE 传送到 #oTLYel
   IF #TPPB.LampTest OR "DB1000_StdSignal".LampTest THEN
       #oTLYel := TRUE;
   END_IF;
   // 含义：条件 #TPPB.LampTest OR "DB1000_StdSignal".LampTest 成立时，将 TRUE 传送到 #oTLGreen
   IF #TPPB.LampTest OR "DB1000_StdSignal".LampTest THEN
       #oTLGreen := TRUE;
   END_IF;
   // 含义：条件 #TPPB.LampTest OR "DB1000_StdSignal".LampTest 成立时，将 TRUE 传送到 #oPanelG
   IF #TPPB.LampTest OR "DB1000_StdSignal".LampTest THEN
       #oPanelG := TRUE;
   END_IF;
   // 含义：条件 #TPPB.LampTest OR "DB1000_StdSignal".LampTest 成立时，将 TRUE 传送到 #oPanelRed
   IF #TPPB.LampTest OR "DB1000_StdSignal".LampTest THEN
       #oPanelRed := TRUE;
   END_IF;
   // 含义：条件 #TPPB.LampTest OR "DB1000_StdSignal".LampTest 成立时，将 TRUE 传送到 #oBeeper
   IF #TPPB.LampTest OR "DB1000_StdSignal".LampTest THEN
       #oBeeper := TRUE;
   END_IF;
   // 含义：条件 #TPPB.LampTest OR "DB1000_StdSignal".LampTest 成立时，将 TRUE 传送到 #oTLBlue
   IF #TPPB.LampTest OR "DB1000_StdSignal".LampTest THEN
       #oTLBlue := TRUE;
   END_IF;
   // 含义：条件 #TPPB.LampTest OR "DB1000_StdSignal".LampTest 成立时，将 TRUE 传送到 #OUT.oPanelHome
   IF #TPPB.LampTest OR "DB1000_StdSignal".LampTest THEN
       #OUT.oPanelHome := TRUE;
   END_IF;

   // ---------- 网络 25 ----------
   // 标题：日光灯控制
   // 含义：当 #TPPB.LampCtrol 为 TRUE 时置位 #oLightingLampClose，否则复位（触点→线圈）
   IF #TPPB.LampCtrol THEN
       #oLightingLampClose := TRUE;
   ELSE
       #oLightingLampClose := FALSE;
   END_IF;

   // ---------- 网络 26 ----------
   // 标题：设备进入特殊模式信息提示
   // 含义：当 #TPPB.EmptyMode 为 TRUE 时置位 #oEmptyMode，否则复位（触点→线圈）
   IF #TPPB.EmptyMode THEN
       #oEmptyMode := TRUE;
   ELSE
       #oEmptyMode := FALSE;
   END_IF;
   // 含义：当 #TPPB.StepMode 为 TRUE 时置位 #oStepMode，否则复位（触点→线圈）
   IF #TPPB.StepMode THEN
       #oStepMode := TRUE;
   ELSE
       #oStepMode := FALSE;
   END_IF;

   // ---------- 网络 27 ----------
   // 标题：单步按钮
   // 含义：条件 "DB1000_StdSignal".PLS.InitialPls 成立时，将 0 传送到 #AtTPPB
   IF "DB1000_StdSignal".PLS.InitialPls THEN
       #AtTPPB := 0;
   END_IF;

   // ---------- 网络 28 ----------
   // （空白网络）
END_FUNCTION_BLOCK

FUNCTION_BLOCK "FB1010_Parameter"   // FB1010, SCL
{ S7_Optimized_Access := 'TRUE' }
// ============================================================
//  Block: FB1010_Parameter
//  ============================================================
//  编号：FB1010
//  原始语言：SCL（规则翻译为 SCL）
//  含义：由 LAD/FBD 网络折叠生成的等效 SCL，导入前请人工复核
   VAR_INPUT
      IMaxProgNo : Int := 300;   // 最大能存储的程序号数量
   END_VAR
   VAR
      TP_Cmd : Word;   // 静态变量
      TP_Status : Word;   // 静态变量
      CmdAuto : Struct   // //触摸屏命令
         ParaSave : Bool;   // 参数保存按钮；
         TypeConfirm : Bool;   // 换型确认按钮
         ParaRead : Bool;   // 请求重新载入参数到编辑区
         ParaCopy : Bool;   // 复制程序号，除了名称
         CopyDestTypeNameSave : Bool;   // 复制目标名称保存
         CopyDestTypeNameRead : Bool;   // 读取复制目标的名称
      END_STRUCT;
      ATCmdAuto : Word;   // 静态变量
      CmdMid : Struct   // 静态变量
         ParaSave : Bool;   // 参数保存按钮；
         TypeConfirm : Bool;   // 换型确认按钮
         ParaRead : Bool;   // 请求重新载入参数到编辑区
         ParaCopy : Bool;   // 复制程序号，除了名称
         CopyDestTypeNameSave : Bool;   // 复制目标名称保存
         CopyDestTypeNameRead : Bool;   // 读取复制目标的名称
      END_STRUCT;
      AtCmdMid_word : Word;   // 静态变量
      Status : Struct   // //触摸屏指示灯
         Para_Saved : Bool;   // 用于确认触摸屏按钮被按下
         TypeChangeConfirmed : Bool;   // On表示确认成功；
         Para_ReNewEdPls : Bool;   // On表示参数发生了更新；
         ParaReadOK : Bool;   // 静态变量
         DBLProcessErr : Bool;   // LoadMemory Process Fail !
         xp3 : Bool;   // 静态变量
         xp4 : Bool;   // 静态变量
         xp5 : Bool;   // 静态变量
         ProgNOEChangeLimit1 : Bool;   // 选型- 键翻页到头
         ProgNOEChangeLimit2 : Bool;   // 选型 + 键翻页到头
         ProgNOCopyDestLimit3 : Bool;   // 静态变量
         ResetParaSaved_DT : Bool;   // 静态变量
      END_STRUCT;
      AtStatus : Word;   // 静态变量
      CurProgNoE : Int := 1;   // 当前程序号编辑区；
      CurProgNoR : Int := 1;   // 当前程序号运行区；
      ProgNoCopyDest : Int := 1;   // 程序选择页面显示的起始编号；
      Aux : Struct   // 静态变量
         AuxTypePara : "UDT_TypePara";   // 静态变量
         CurProgNoEBake : Int := 0;   // 用于指定要拷贝的程序号目的地
         ProgNoCopyDest_Bake : Int := 1;   // 程序选择页面显示的起始编号；
         ReadTypeNameIndex : Int;   // 从1开始
         CurProgNO_Ten_E : Int;   // CurProtNOE的10位数
         CurProgNO_Ten_E_Bake : Int := -100;   // 静态变量
         DefaultTypePara : "UDT_TypePara";   // 静态变量
         ReadTypeParaDBL : Struct   // 676
            Cmd : Bool;   // 数据尚未从装载存储器读取
            CmdReqPls : Bool;   // 静态变量
            Busy : Bool;   // 静态变量
            Index : Int;   // 静态变量
            Read_DBL_RetVal : Int;   // 静态变量
         END_STRUCT;
         WriteTypeParaDBL : Struct   // 静态变量
            Cmd : Bool;   // 静态变量
            CmdReqPls : Bool;   // 静态变量
            Busy : Bool;   // 静态变量
            Index : Int;   // 静态变量
            Write_DBL_RetVal : Int;   // 静态变量
         END_STRUCT;
         ReadSystemParaDBL : Struct   // 676
            Cmd : Bool;   // 数据尚未从装载存储器读取
            CmdReqPls : Bool;   // 静态变量
            Busy : Bool;   // 静态变量
            Index : Int;   // 静态变量
            Read_DBL_RetVal : Int;   // 静态变量
         END_STRUCT;
         WriteSystemParaDBL : Struct   // 静态变量
            Cmd : Bool;   // 静态变量
            CmdReqPls : Bool;   // 静态变量
            Busy : Bool;   // 静态变量
            Index : Int;   // 静态变量
            Write_DBL_RetVal : Int;   // 静态变量
         END_STRUCT;
      END_STRUCT;
      "step" : Int;   // 静态变量
      AryTypeName : Array[1..11] of String[20];   // 产品型号选择页面显示的产品名称；
      At_TypeName : Array[22..263] of Byte;   // 静态变量
      ArrayProgNoForSel : Array[1..10] of Int;   // 静态变量
      SystemParaE : "UDT_SystemPara";   // 系统参数_编辑区280
      SystemParaR : "UDT_SystemPara";   // 系统参数_运行区480
      TypeParaE : "UDT_TypePara";   // 产品参数_编辑区680
      AtTypeParaETypeName : Byte;   // 静态变量
      TypeParaR : "UDT_TypePara";   // 产品参数_运行区776
      TypeName : String[20];   // 静态变量
      bit : Struct   // 静态变量
         Bit0 : Bool;   // 静态变量
         sp : Word;   // 静态变量
         Other : Struct   // 静态变量
            Bool_1 : Bool;   // 静态变量
            Byte_2 : Byte;   // 静态变量
            Int_1 : Int;   // 静态变量
            "Char" : Char;   // 静态变量
         END_STRUCT;
      END_STRUCT;
      Other : Struct   // 静态变量
         STxxxCCDProgNO : Int;   // 静态变量
         FixtureEnable : Bool;   // 静态变量
         Byte_1 : Byte;   // 静态变量
         Int_1 : Int;   // 静态变量
         "Char" : Char;   // 静态变量
         Word_1 : Word;   // 静态变量
         DInt_1 : DInt;   // 静态变量
         DWord_1 : DWord;   // 静态变量
         Real_1 : Real;   // 静态变量
         S5Time : Time;   // 静态变量
         "String" : String[5];   // 静态变量
      END_STRUCT;
   END_VAR
   VAR_TEMP
      index : Int;   // 临时变量
      T_CurProgNO_E : Int;   // 临时变量
   END_VAR
BEGIN

   // ---------- 网络 1 ----------
   // 含义：本网络为 StructuredText（SCL）原文重建，非 LAD 折叠
   IF #step = 0
   THEN
       #AtCmdMid_word := #ATCmdAuto OR #TP_Cmd;
       #TP_Cmd := 0;
       #ATCmdAuto := 0;
       IF (#ProgNoCopyDest <> #Aux.ProgNoCopyDest_Bake) THEN
           #CmdAuto.CopyDestTypeNameRead := TRUE;
           #Aux.ProgNoCopyDest_Bake := #ProgNoCopyDest;
       END_IF;
       IF (#CurProgNoE <> #Aux.CurProgNoEBake) THEN
           #step := 1999;
           #Aux.CurProgNoEBake := #CurProgNoE;
       END_IF;
       IF #AtCmdMid_word <> 0 THEN
           #step := (ENCO(IN := #AtCmdMid_word) - 8 + 1) * 100;
       END_IF;
       IF "DB1000_StdSignal".PLS.PS10 AND #Status.Para_Saved THEN
           IF #Status.ResetParaSaved_DT = TRUE THEN
               #Status.ResetParaSaved_DT := FALSE;
               #Status.Para_Saved := FALSE;
           ELSE
               #Status.ResetParaSaved_DT := TRUE;
           END_IF;
       END_IF;
   END_IF;
   #TP_Status := #AtStatus;
   #Status.Para_ReNewEdPls := FALSE;
   #Status.TypeChangeConfirmed := (#CurProgNoR = #CurProgNoE);
   #Status.ProgNOEChangeLimit1 := (#CurProgNoE >= #IMaxProgNo);
   #Status.ProgNOEChangeLimit2 := (#CurProgNoE > (#IMaxProgNo - 10));
   #Status.ProgNOCopyDestLimit3 := (#ProgNoCopyDest >= #IMaxProgNo);
   IF (#Aux.WriteTypeParaDBL.Cmd = TRUE)
   THEN
       #Aux.WriteTypeParaDBL.Write_DBL_RetVal := WRIT_DBL(REQ := #Aux.WriteTypeParaDBL.CmdReqPls,
                                                          SRCBLK := #Aux.AuxTypePara,
                                                          BUSY => #Aux.WriteTypeParaDBL.Busy,
                                                          DSTBLK => "DB5000_ParameterLoadMemory".AryTypePara[#Aux.WriteTypeParaDBL.Index]);
       IF (#Aux.WriteTypeParaDBL.Busy)
       THEN
           #Aux.WriteTypeParaDBL.CmdReqPls := FALSE;
           RETURN;
       END_IF;
       IF (#Aux.WriteTypeParaDBL.Busy = FALSE)
       THEN
           #Aux.WriteTypeParaDBL.Cmd := FALSE;
           IF (#Aux.WriteTypeParaDBL.Write_DBL_RetVal <> 0)
           THEN
               #Status.DBLProcessErr := TRUE;
               #step := 0;
           ELSE
               #Status.DBLProcessErr := FALSE;
           END_IF;
       END_IF;
   END_IF;
   IF (#Aux.ReadTypeParaDBL.Cmd) THEN
       #Aux.ReadTypeParaDBL.Read_DBL_RetVal := READ_DBL(REQ := #Aux.ReadTypeParaDBL.CmdReqPls,
                                                        SRCBLK := "DB5000_ParameterLoadMemory".AryTypePara[#Aux.ReadTypeParaDBL.Index],
                                                        BUSY => #Aux.ReadTypeParaDBL.Busy,
                                                        DSTBLK => #Aux.AuxTypePara);
       IF (#Aux.ReadTypeParaDBL.Busy = TRUE)
       THEN
           #Aux.ReadTypeParaDBL.CmdReqPls := FALSE;
           RETURN;
       END_IF;
       IF (#Aux.ReadTypeParaDBL.Busy = FALSE)
       THEN
           #Aux.ReadTypeParaDBL.Cmd := FALSE;
           IF (#Aux.ReadTypeParaDBL.Read_DBL_RetVal <> 0)
           THEN
               #Status.DBLProcessErr := TRUE;
               #step := 0;
           ELSE
               #Status.DBLProcessErr := FALSE;
           END_IF;
       END_IF;
   END_IF;
   IF (#Aux.WriteSystemParaDBL.Cmd = TRUE)
   THEN
       #Aux.WriteSystemParaDBL.Write_DBL_RetVal := WRIT_DBL(REQ := #Aux.WriteSystemParaDBL.CmdReqPls,
                                                            SRCBLK := #SystemParaE,
                                                            BUSY => #Aux.WriteSystemParaDBL.Busy,
                                                            DSTBLK => "DB5000_ParameterLoadMemory".SystemParaE);
       IF (#Aux.WriteSystemParaDBL.Busy)
       THEN
           #Aux.WriteSystemParaDBL.CmdReqPls := FALSE;
           RETURN;
       END_IF;
       IF (#Aux.WriteSystemParaDBL.Busy = FALSE)
       THEN
           #Aux.WriteSystemParaDBL.Cmd := FALSE;
           IF (#Aux.WriteSystemParaDBL.Write_DBL_RetVal <> 0)
           THEN
               #Status.DBLProcessErr := TRUE;
               #step := 0;
           ELSE
               #SystemParaR := #SystemParaE;
               #Status.DBLProcessErr := FALSE;
           END_IF;
       END_IF;
   END_IF;
   IF (#Aux.ReadSystemParaDBL.Cmd) THEN
       #Aux.ReadSystemParaDBL.Read_DBL_RetVal := READ_DBL(REQ := #Aux.ReadSystemParaDBL.CmdReqPls,
                                                          SRCBLK := "DB5000_ParameterLoadMemory".SystemParaE,
                                                          BUSY => #Aux.ReadSystemParaDBL.Busy,
                                                          DSTBLK => #SystemParaE);
       IF (#Aux.ReadSystemParaDBL.Busy = TRUE)
       THEN
           #Aux.ReadSystemParaDBL.CmdReqPls := FALSE;
           RETURN;
       END_IF;
       IF (#Aux.ReadSystemParaDBL.Busy = FALSE)
       THEN
           #Aux.ReadSystemParaDBL.Cmd := FALSE;
           IF (#Aux.ReadSystemParaDBL.Read_DBL_RetVal <> 0)
           THEN
               #Status.DBLProcessErr := TRUE;
               #step := 0;
           ELSE
               #Status.DBLProcessErr := FALSE;
               #SystemParaR := #SystemParaE;
           END_IF;
       END_IF;
   END_IF;
   CASE #step OF
       100:
           #AtTypeParaETypeName := 20;
           #Aux.AuxTypePara := #TypeParaE;
           #Aux.WriteTypeParaDBL.Index := #CurProgNoE;
           #step := #step + 1;
           #Aux.WriteSystemParaDBL.Cmd := TRUE;
           #Aux.WriteSystemParaDBL.CmdReqPls := true;
       200, 400:
           #Aux.ReadTypeParaDBL.Index := #CurProgNoE;
           #step := #step + 1;
       300:
           #CurProgNoE := #CurProgNoR;
           #Aux.ReadTypeParaDBL.Index := #CurProgNoE;
           #step := #step + 1;
           #Aux.ReadSystemParaDBL.Cmd := TRUE;
           #Aux.ReadSystemParaDBL.CmdReqPls := true;
       500, 600:
           #Aux.ReadTypeParaDBL.Index := #ProgNoCopyDest;
           #step := #step + 1;
       1999:
           #Aux.CurProgNO_Ten_E := (#CurProgNoE - 1) - (#CurProgNoE - 1) MOD 10;
           #Aux.ReadTypeNameIndex := 1;
           IF (#Aux.CurProgNO_Ten_E = #Aux.CurProgNO_Ten_E_Bake)
           THEN
               #Aux.ReadTypeParaDBL.Index := #CurProgNoE;
               #step := 301;
           ELSE
               #step := #step + 1;
           END_IF;
       2000:
           #Aux.ReadTypeParaDBL.Index := #Aux.CurProgNO_Ten_E + #Aux.ReadTypeNameIndex;
           #step := #step + 1;
       101:
           #Aux.WriteTypeParaDBL.Cmd := TRUE;
           #Aux.WriteTypeParaDBL.CmdReqPls := true;
           #step := #step + 1;
       201, 301, 401, 501, 601, 2001:
           #Aux.ReadTypeParaDBL.Cmd := TRUE;
           #Aux.ReadTypeParaDBL.CmdReqPls := TRUE;
           #step := #step + 1;
       102, 202, 302, 402, 502, 602, 2002:
           IF (#Aux.WriteTypeParaDBL.Cmd = FALSE)
               AND (#Aux.ReadTypeParaDBL.Cmd = FALSE)
               AND (#Aux.WriteSystemParaDBL.Cmd = false)
               AND (#Aux.ReadSystemParaDBL.Cmd = false)
           THEN
               #step := #step + 8;
           END_IF;
       110:
           IF #CurProgNoE = #CurProgNoR THEN
               #TypeParaR := #TypeParaE;
               #Status.Para_ReNewEdPls := TRUE;
           END_IF;
           #Status.Para_Saved := TRUE;
           #SystemParaR := #SystemParaE;
           #step := 1999;
       210:
           #CurProgNoR := #CurProgNoE;
           #TypeParaE := #Aux.AuxTypePara;
           #TypeParaR := #TypeParaE;
           #Status.Para_ReNewEdPls := TRUE;
           #step := 0;
       310:
           #TypeParaE := #Aux.AuxTypePara;
           #SystemParaE := #SystemParaR;
           #step := 0;
       410:
           #Aux.AuxTypePara := #TypeParaE;
           #Aux.AuxTypePara.TypeName := 'new,NoName';
           #AryTypeName[11] := #Aux.AuxTypePara.TypeName;
           #Aux.WriteTypeParaDBL.Cmd := TRUE;
           #Aux.WriteTypeParaDBL.CmdReqPls := TRUE;
           #Aux.WriteTypeParaDBL.Index := #ProgNoCopyDest;
           #step := 0;
       510:
           #Aux.AuxTypePara.TypeName := #AryTypeName[11];
           #Aux.WriteTypeParaDBL.Cmd := TRUE;
           #Aux.WriteTypeParaDBL.CmdReqPls := TRUE;
           #Aux.WriteTypeParaDBL.Index := #ProgNoCopyDest;
           #step := 0;
       610:
           #AryTypeName[11] := #Aux.AuxTypePara.TypeName;
           #step := 0;
       2010:
           #At_TypeName[#Aux.ReadTypeNameIndex] := 20;
           #AryTypeName[#Aux.ReadTypeNameIndex] := #Aux.AuxTypePara.TypeName;
           #ArrayProgNoForSel[#Aux.ReadTypeNameIndex] := #Aux.ReadTypeParaDBL.Index;
           IF (#Aux.ReadTypeParaDBL.Index = 1) THEN
               #Aux.DefaultTypePara := #Aux.AuxTypePara;
           END_IF;
           #Aux.ReadTypeNameIndex := #Aux.ReadTypeNameIndex + 1;
           IF #CurProgNoE = #Aux.ReadTypeParaDBL.Index THEN
               #TypeParaE := #Aux.AuxTypePara;
           END_IF;
           IF #Aux.ReadTypeNameIndex <= 10 THEN
               #step := 2000;
           ELSE
               #step := 2020;
           END_IF;
       2020:
           IF #TypeParaE.TypeName = '' THEN
               #TypeParaE := #Aux.DefaultTypePara;
               #TypeParaE.TypeName := '';
           END_IF;
           #Aux.CurProgNO_Ten_E_Bake := #Aux.CurProgNO_Ten_E;
           #step := 0;
       ELSE:
           #step := 0;
   END_CASE;
END_FUNCTION_BLOCK

FUNCTION_BLOCK "FB1089_AddrRegister"   // FB1089, SCL
{ S7_Optimized_Access := 'TRUE' }
// ============================================================
//  Block: FB1089_AddrRegister
//  ============================================================
//  编号：FB1089
//  原始语言：SCL（规则翻译为 SCL）
//  含义：由 LAD/FBD 网络折叠生成的等效 SCL，导入前请人工复核
   VAR
      Siemens_V90_Servo_V3 : Struct   // Siemens V90 伺服偏移地址处理；
         FBCall_StartAddr : Int;   // FB块被调用的起始地址
         FBCall_IndexNO : Int := 1;   // FB块数组被调用的编号，从1开始，0无效
         FB_ByteLength : Int := 800;   // FB块调用时所占的地址长度
         Aux : Struct   // 静态变量
            FBCall_StartAddr : Int;   // FB块被调用的起始地址
            FBCall_IndexNO : Int;   // FB块数组被调用的编号，从1开始，0无效
            StartAddr : Int;   // 静态变量
         END_STRUCT;
         TotalRunnningDistance : Int;   // 静态变量
         TP_Cmd : Int;   // 静态变量
         TP_Status : Int;   // 静态变量
         CTRL_IN_SetValueVelocity : Int;   // 静态变量
         CTRL_IN_SetValuePosition : Int;   // 静态变量
         CTRL_IN_SetValueTorque : Int;   // 静态变量
         CTRL_IN_PNU : Int;   // 静态变量
         CTRL_IN_ParameterValue_DataCom : Int;   // 静态变量
         CTRL_IN_InitParameter_Min_SetValuePosition : Int;   // 静态变量
         CTRL_IN_InitParameter_Max_SetValuePosition : Int;   // 静态变量
         CTRL_IN_TraversingBlockNO : Int;   // 静态变量
         CTRL_OUT_ActualPosition : Int;   // 静态变量
         CTRL_OUT_ActualVelocity : Int;   // 静态变量
         CTRL_OUT_ParameterValue_DataCom : Int;   // 静态变量
         CTRL_OUT_MotorRatedTorque : Int;   // 静态变量
         CTRL_OUT_LastCylceTime : Int;   // 静态变量
         CTRL_OUT_Max_SetValueVelocity : Int;   // 静态变量
         Status_PromptValue : Int;   // 静态变量
         Bus_IN_Data_Fault_Code : Int;   // 静态变量
      END_STRUCT;
      Festo_Servo_V1 : Struct   // Festo 伺服偏移地址处理；
         FBCall_StartAddr : Int;   // FB块被调用的起始地址
         FBCall_IndexNO : Int := 1;   // FB块数组被调用的编号，从1开始，0无效
         FB_ByteLength : Int := 800;   // FB块调用时所占的地址长度
         Aux : Struct   // 静态变量
            FBCall_StartAddr : Int;   // FB块被调用的起始地址
            FBCall_IndexNO : Int;   // FB块数组被调用的编号，从1开始，0无效
            StartAddr : Int;   // 静态变量
         END_STRUCT;
         TotalRunnningDistance : Int;   // 静态变量
         TP_Cmd : Int;   // 静态变量
         TP_Status : Int;   // 静态变量
         CTRL_IN_SetValueVelocity : Int;   // 静态变量
         CTRL_IN_SetValuePosition : Int;   // 静态变量
         CTRL_IN_TorqueModeStartRamp : Int;   // 静态变量
         CTRL_IN_SetValueTorque : Int;   // 静态变量
         CTRL_IN_PNU : Int;   // 静态变量
         CTRL_IN_InitParameter_BaseVelocity : Int;   // 静态变量
         CTRL_OUT_ActualPosition : Int;   // 静态变量
         CTRL_OUT_ActualVelocity : Int;   // 静态变量
         CTRL_OUT_MotorRatedTorque : Int;   // 静态变量
         CTRL_OUT_LastCylceTime : Int;   // 静态变量
         Status_PromptValue : Int;   // 静态变量
      END_STRUCT;
      TCPIP_Client_V3 : Struct   // TCPIP_Client偏移地址处理；
         FB_ByteLength : Int := 1000;   // FB块调用时所占的地址长度
         FBCall_StartAddr : Int;   // FB块被调用的起始地址
         FBCall_IndexNO : Int := 1;   // FB块数组被调用的编号，从1开始，0无效
         Aux : Struct   // 静态变量
            FBCall_StartAddr : Int;   // FB块被调用的起始地址
            FBCall_IndexNO : Int;   // FB块数组被调用的编号，从1开始，0无效
            StartAddr : Int;   // 静态变量
         END_STRUCT;
         TP_Cmd : Int;   // 静态变量
         TP_Status : Int;   // 静态变量
         Ctrl_IN_TCPIP_ServerIP_High : Int;   // 静态变量
         Ctrl_IN_TCPIP_ServerIP_Mid1 : Int;   // 静态变量
         Ctrl_IN_TCPIP_ServerIP_Mid2 : Int;   // 静态变量
         Ctrl_IN_TCPIP_ServerIP_Low : Int;   // 静态变量
         Ctrl_IN_TCPIP_ServerPort : Int;   // 静态变量
         Ctrl_IN_SendStr : Int;   // 静态变量
         Ctrl_Out_RecvStr : Int;   // 静态变量
         Ctrl_Out_TCPIP_Recv_Status : Int;   // 静态变量
         Ctrl_Out_LastCylceTime : Int;   // 静态变量
         Status_PromptValue : Int;   // 静态变量
      END_STRUCT;
      Congex_InsightCCD_V1 : Struct   // Congex_InsightCCD偏移地址处理；
         FBCall_StartAddr : Int;   // FB块被调用的起始地址
         FBCall_IndexNO : Int := 1;   // FB块数组被调用的编号，从1开始，0无效
         FB_ByteLength : Int := 300;   // FB块调用时所占的地址长度
         Aux : Struct   // 静态变量
            FBCall_StartAddr : Int;   // FB块被调用的起始地址
            FBCall_IndexNO : Int;   // FB块数组被调用的编号，从1开始，0无效
            StartAddr : Int;   // 静态变量
         END_STRUCT;
         TP_Cmd : Int;   // 静态变量
         TP_Status : Int;   // 静态变量
         CTRL_IN_ProgNo : Int;   // 静态变量
         CTRL_OUT_OKCounter : Int;   // 静态变量
         CTRL_OUT_NOKCounter : Int;   // 静态变量
         OUT_LastCylceTime : Int;   // 静态变量
         Status_PromptValue : Int;   // 静态变量
      END_STRUCT;
      AteqLeakTest_TCP2RS232ModBus_V1 : Struct   // Ateq偏移地址处理；
         FBCall_StartAddr : Int;   // FB块被调用的起始地址
         FBCall_IndexNO : Int := 1;   // FB块数组被调用的编号，从1开始，0无效
         FB_ByteLength : Int := 1800;   // FB块调用时所占的地址长度
         Aux : Struct   // 静态变量
            FBCall_StartAddr : Int;   // FB块被调用的起始地址
            FBCall_IndexNO : Int;   // FB块数组被调用的编号，从1开始，0无效
            StartAddr : Int;   // 静态变量
         END_STRUCT;
         TP_Cmd : Int;   // 静态变量
         TP_Status : Int;   // 静态变量
         CTRL_IN_ProgNo : Int;   // 静态变量
         Ctrl_IN_ModBusSlaveNO : Int;   // 静态变量
         CTRL_Out_ProgNo : Int;   // 静态变量
         CTRL_OUT_OKCounter : Int;   // 静态变量
         CTRL_OUT_NOKCounter : Int;   // 静态变量
         CTRL_OUT_LastCylceTime : Int;   // 静态变量
         CTRL_OUT_Pressure : Int;   // 静态变量
         CTRL_OUT_LeakRate : Int;   // 静态变量
         Status_PromptValue : Int;   // 静态变量
      END_STRUCT;
      IFM_O2D22X_TCP_V1 : Struct   // IFM O2D22x轮廓传感器地址处理
         FBCall_StartAddr : Int;   // FB块被调用的起始地址
         FBCall_IndexNO : Int := 1;   // FB块数组被调用的编号，从1开始，0无效
         FB_ByteLength : Int := 1300;   // FB块调用时所占的地址长度
         Aux : Struct   // 静态变量
            FBCall_StartAddr : Int;   // FB块被调用的起始地址
            FBCall_IndexNO : Int;   // FB块数组被调用的编号，从1开始，0无效
            StartAddr : Int;   // 静态变量
         END_STRUCT;
         TP_Cmd : Int;   // 静态变量
         TP_Status : Int;   // 静态变量
         CTRL_IN_ProgNo : Int;   // 静态变量
         CTRL_IN_DigitOutPutsOKBit : Int;   // 静态变量
         CTRL_Out_ProgNo : Int;   // 静态变量
         CTRL_OUT_OKCounter : Int;   // 静态变量
         CTRL_OUT_NOKCounter : Int;   // 静态变量
         CTRL_OUT_LastCylceTime : Int;   // 静态变量
         CTRL_OUT_DigitOutPutsOKBit : Int;   // 静态变量
         Status_PromptValue : Int;   // 静态变量
      END_STRUCT;
      BisArrayInfo_V4 : Struct   // Balluff_RFID_调用数组信息
         TP_Bis_Index : Int := 1;   // 触摸屏使用，从1~开始
         TP_Bis_Index_Max : Int := 1;   // 人工输入
         TP_BisDataStructLength : Int := 100;   // 静态变量
         TP_BisArrayStartAddress : Int;   // 静态变量
      END_STRUCT;
      Analog_IN_V4 : Struct   // AI_模拟量输入处理
         FBCall_StartAddr : Int;   // FB块被调用的起始地址
         FBCall_IndexNO : Int := 1;   // FB块数组被调用的编号，从1开始，0无效
         FB_ByteLength : Int := 200;   // FB块调用时所占的地址长度
         Aux : Struct   // 静态变量
            FBCall_StartAddr : Int;   // FB块被调用的起始地址
            FBCall_IndexNO : Int;   // FB块数组被调用的编号，从1开始，0无效
            StartAddr : Int;   // 静态变量
         END_STRUCT;
         TP_Cmd : Int;   // 静态变量
         CTRL_IN_TP_AI_Gain : Int;   // 静态变量
         CTRL_IN_TP_AI_OffSet : Int;   // 静态变量
         CTRL_IN_TP_PreSetValue : Int;   // 静态变量
         CTRL_IN_TP_ActualAI_1 : Int;   // 静态变量
         CTRL_IN_TP_ActualAI_2 : Int;   // 静态变量
         CTRL_IN_TP_ActualAI_Value1 : Int;   // 静态变量
         CTRL_IN_TP_ActualAI_Value2 : Int;   // 静态变量
         CTRL_OUT_Cur_Val_Out : Int;   // 静态变量
         CTRL_OUT_TrigerValue : Int;   // 静态变量
         CTRL_OUT_TrigerValue_Array : Int;   // 静态变量
         CTRL_OUT_TrigerTPColorStatus_Array : Int;   // 静态变量
         CTRL_OUT_TrigerCounter : Int;   // 静态变量
      END_STRUCT;
   END_VAR
   VAR_TEMP
      T_Index : DInt;   // 临时变量
   END_VAR
BEGIN

   // ---------- 网络 1 ----------
   // 含义：本网络为 StructuredText（SCL）原文重建，非 LAD 折叠
   IF #Siemens_V90_Servo_V3.FBCall_StartAddr <> #Siemens_V90_Servo_V3.Aux.FBCall_StartAddr
       OR #Siemens_V90_Servo_V3.FBCall_IndexNO <> #Siemens_V90_Servo_V3.Aux.FBCall_IndexNO THEN
       #Siemens_V90_Servo_V3.Aux.FBCall_StartAddr := #Siemens_V90_Servo_V3.FBCall_StartAddr;
       #Siemens_V90_Servo_V3.Aux.FBCall_IndexNO := #Siemens_V90_Servo_V3.FBCall_IndexNO;
       #Siemens_V90_Servo_V3.Aux.StartAddr := #Siemens_V90_Servo_V3.Aux.FBCall_StartAddr +
       (#Siemens_V90_Servo_V3.Aux.FBCall_IndexNO - 1) *
       #Siemens_V90_Servo_V3.FB_ByteLength;
       #Siemens_V90_Servo_V3.TotalRunnningDistance := #Siemens_V90_Servo_V3.Aux.StartAddr + 8;
       #Siemens_V90_Servo_V3.TP_Cmd := #Siemens_V90_Servo_V3.Aux.StartAddr + 12;
       #Siemens_V90_Servo_V3.TP_Status := #Siemens_V90_Servo_V3.Aux.StartAddr + 14;
       #Siemens_V90_Servo_V3.CTRL_IN_SetValueVelocity := #Siemens_V90_Servo_V3.Aux.StartAddr + 20;
       #Siemens_V90_Servo_V3.CTRL_IN_SetValuePosition := #Siemens_V90_Servo_V3.Aux.StartAddr + 24;
       #Siemens_V90_Servo_V3.CTRL_IN_SetValueTorque := #Siemens_V90_Servo_V3.Aux.StartAddr + 32;
       #Siemens_V90_Servo_V3.CTRL_IN_TraversingBlockNO := #Siemens_V90_Servo_V3.Aux.StartAddr + 36;
       #Siemens_V90_Servo_V3.CTRL_IN_PNU := #Siemens_V90_Servo_V3.Aux.StartAddr + 42;
       #Siemens_V90_Servo_V3.CTRL_IN_ParameterValue_DataCom := #Siemens_V90_Servo_V3.Aux.StartAddr + 46;
       #Siemens_V90_Servo_V3.CTRL_IN_InitParameter_Min_SetValuePosition := #Siemens_V90_Servo_V3.Aux.StartAddr + 64;
       #Siemens_V90_Servo_V3.CTRL_IN_InitParameter_Max_SetValuePosition := #Siemens_V90_Servo_V3.Aux.StartAddr + 68;
       #Siemens_V90_Servo_V3.CTRL_OUT_ActualPosition := #Siemens_V90_Servo_V3.Aux.StartAddr + 160;
       #Siemens_V90_Servo_V3.CTRL_OUT_ActualVelocity := #Siemens_V90_Servo_V3.Aux.StartAddr + 164;
       #Siemens_V90_Servo_V3.CTRL_OUT_ParameterValue_DataCom := #Siemens_V90_Servo_V3.Aux.StartAddr + 168;
       #Siemens_V90_Servo_V3.CTRL_OUT_MotorRatedTorque := #Siemens_V90_Servo_V3.Aux.StartAddr + 172;
       #Siemens_V90_Servo_V3.CTRL_OUT_LastCylceTime := #Siemens_V90_Servo_V3.Aux.StartAddr + 176;
       #Siemens_V90_Servo_V3.CTRL_OUT_Max_SetValueVelocity := #Siemens_V90_Servo_V3.Aux.StartAddr + 180;
       #Siemens_V90_Servo_V3.Status_PromptValue := #Siemens_V90_Servo_V3.Aux.StartAddr + 206;
       #Siemens_V90_Servo_V3.Bus_IN_Data_Fault_Code := #Siemens_V90_Servo_V3.Aux.StartAddr + 228;
   END_IF;
   IF #Festo_Servo_V1.FBCall_StartAddr <> #Festo_Servo_V1.Aux.FBCall_StartAddr
       OR #Festo_Servo_V1.FBCall_IndexNO <> #Festo_Servo_V1.Aux.FBCall_IndexNO THEN
       #Festo_Servo_V1.Aux.FBCall_StartAddr := #Festo_Servo_V1.FBCall_StartAddr;
       #Festo_Servo_V1.Aux.FBCall_IndexNO := #Festo_Servo_V1.FBCall_IndexNO;
       #Festo_Servo_V1.Aux.StartAddr := #Festo_Servo_V1.Aux.FBCall_StartAddr +
       (#Festo_Servo_V1.Aux.FBCall_IndexNO - 1) *
       #Festo_Servo_V1.FB_ByteLength;
       #Festo_Servo_V1.TotalRunnningDistance := #Festo_Servo_V1.Aux.StartAddr + 18;
       #Festo_Servo_V1.TP_Cmd := #Festo_Servo_V1.Aux.StartAddr + 22;
       #Festo_Servo_V1.TP_Status := #Festo_Servo_V1.Aux.StartAddr + 24;
       #Festo_Servo_V1.CTRL_IN_SetValueVelocity := #Festo_Servo_V1.Aux.StartAddr + 30;
       #Festo_Servo_V1.CTRL_IN_SetValuePosition := #Festo_Servo_V1.Aux.StartAddr + 34;
       #Festo_Servo_V1.CTRL_IN_TorqueModeStartRamp := #Festo_Servo_V1.Aux.StartAddr + 38;
       #Festo_Servo_V1.CTRL_IN_SetValueTorque := #Festo_Servo_V1.Aux.StartAddr + 42;
       #Festo_Servo_V1.CTRL_IN_PNU := #Festo_Servo_V1.Aux.StartAddr + 46;
       #Festo_Servo_V1.CTRL_IN_InitParameter_BaseVelocity := #Festo_Servo_V1.Aux.StartAddr + 58;
       #Festo_Servo_V1.CTRL_OUT_ActualPosition := #Festo_Servo_V1.Aux.StartAddr + 78;
       #Festo_Servo_V1.CTRL_OUT_ActualVelocity := #Festo_Servo_V1.Aux.StartAddr + 82;
       #Festo_Servo_V1.CTRL_OUT_MotorRatedTorque := #Festo_Servo_V1.Aux.StartAddr + 84;
       #Festo_Servo_V1.CTRL_OUT_LastCylceTime := #Festo_Servo_V1.Aux.StartAddr + 88;
       #Festo_Servo_V1.Status_PromptValue := #Festo_Servo_V1.Aux.StartAddr + 102;
   END_IF;
   IF #TCPIP_Client_V3.FBCall_StartAddr <> #TCPIP_Client_V3.Aux.FBCall_StartAddr
       OR #TCPIP_Client_V3.FBCall_IndexNO <> #TCPIP_Client_V3.Aux.FBCall_IndexNO THEN
       #TCPIP_Client_V3.Aux.FBCall_StartAddr := #TCPIP_Client_V3.FBCall_StartAddr;
       #TCPIP_Client_V3.Aux.FBCall_IndexNO := #TCPIP_Client_V3.FBCall_IndexNO;
       #TCPIP_Client_V3.Aux.StartAddr := #TCPIP_Client_V3.Aux.FBCall_StartAddr +
       (#TCPIP_Client_V3.Aux.FBCall_IndexNO - 1) *
       #TCPIP_Client_V3.FB_ByteLength;
       #TCPIP_Client_V3.TP_Cmd := #TCPIP_Client_V3.Aux.StartAddr + 4;
       #TCPIP_Client_V3.TP_Status := #TCPIP_Client_V3.Aux.StartAddr + 8;
       #TCPIP_Client_V3.Ctrl_IN_TCPIP_ServerIP_High := #TCPIP_Client_V3.Aux.StartAddr + 14;
       #TCPIP_Client_V3.Ctrl_IN_TCPIP_ServerIP_Mid1 := #TCPIP_Client_V3.Aux.StartAddr + 15;
       #TCPIP_Client_V3.Ctrl_IN_TCPIP_ServerIP_Mid2 := #TCPIP_Client_V3.Aux.StartAddr + 16;
       #TCPIP_Client_V3.Ctrl_IN_TCPIP_ServerIP_Low := #TCPIP_Client_V3.Aux.StartAddr + 17;
       #TCPIP_Client_V3.Ctrl_IN_TCPIP_ServerPort := #TCPIP_Client_V3.Aux.StartAddr + 18;
       #TCPIP_Client_V3.Ctrl_IN_SendStr := #TCPIP_Client_V3.Aux.StartAddr + 20;
       #TCPIP_Client_V3.Ctrl_Out_RecvStr := #TCPIP_Client_V3.Aux.StartAddr + 312;
       #TCPIP_Client_V3.Ctrl_Out_TCPIP_Recv_Status := #TCPIP_Client_V3.Aux.StartAddr + 568;
       #TCPIP_Client_V3.Ctrl_Out_LastCylceTime := #TCPIP_Client_V3.Aux.StartAddr + 570;
       #TCPIP_Client_V3.Status_PromptValue := #TCPIP_Client_V3.Aux.StartAddr + 576;
   END_IF;
   IF #Congex_InsightCCD_V1.FBCall_StartAddr <> #Congex_InsightCCD_V1.Aux.FBCall_StartAddr
       OR #Congex_InsightCCD_V1.FBCall_IndexNO <> #Congex_InsightCCD_V1.Aux.FBCall_IndexNO THEN
       #Congex_InsightCCD_V1.Aux.FBCall_StartAddr := #Congex_InsightCCD_V1.FBCall_StartAddr;
       #Congex_InsightCCD_V1.Aux.FBCall_IndexNO := #Congex_InsightCCD_V1.FBCall_IndexNO;
       #Congex_InsightCCD_V1.Aux.StartAddr := #Congex_InsightCCD_V1.Aux.FBCall_StartAddr +
       (#Congex_InsightCCD_V1.Aux.FBCall_IndexNO - 1) *
       #Congex_InsightCCD_V1.FB_ByteLength;
       #Congex_InsightCCD_V1.TP_Cmd := #Congex_InsightCCD_V1.Aux.StartAddr + 18;
       #Congex_InsightCCD_V1.TP_Status := #Congex_InsightCCD_V1.Aux.StartAddr + 20;
       #Congex_InsightCCD_V1.CTRL_IN_ProgNo := #Congex_InsightCCD_V1.Aux.StartAddr + 26;
       #Congex_InsightCCD_V1.CTRL_OUT_OKCounter := #Congex_InsightCCD_V1.Aux.StartAddr + 36;
       #Congex_InsightCCD_V1.CTRL_OUT_NOKCounter := #Congex_InsightCCD_V1.Aux.StartAddr + 40;
       #Congex_InsightCCD_V1.OUT_LastCylceTime := #Congex_InsightCCD_V1.Aux.StartAddr + 44;
       #Congex_InsightCCD_V1.Status_PromptValue := #Congex_InsightCCD_V1.Aux.StartAddr + 50;
   END_IF;
   IF #AteqLeakTest_TCP2RS232ModBus_V1.FBCall_StartAddr <> #AteqLeakTest_TCP2RS232ModBus_V1.Aux.FBCall_StartAddr
       OR #AteqLeakTest_TCP2RS232ModBus_V1.FBCall_IndexNO <> #AteqLeakTest_TCP2RS232ModBus_V1.Aux.FBCall_IndexNO THEN
       #AteqLeakTest_TCP2RS232ModBus_V1.Aux.FBCall_StartAddr := #AteqLeakTest_TCP2RS232ModBus_V1.FBCall_StartAddr;
       #AteqLeakTest_TCP2RS232ModBus_V1.Aux.FBCall_IndexNO := #AteqLeakTest_TCP2RS232ModBus_V1.FBCall_IndexNO;
       #AteqLeakTest_TCP2RS232ModBus_V1.Aux.StartAddr := #AteqLeakTest_TCP2RS232ModBus_V1.Aux.FBCall_StartAddr +
       (#AteqLeakTest_TCP2RS232ModBus_V1.Aux.FBCall_IndexNO - 1) *
       #AteqLeakTest_TCP2RS232ModBus_V1.FB_ByteLength;
       #AteqLeakTest_TCP2RS232ModBus_V1.TP_Cmd := #AteqLeakTest_TCP2RS232ModBus_V1.Aux.StartAddr + 4;
       #AteqLeakTest_TCP2RS232ModBus_V1.TP_Status := #AteqLeakTest_TCP2RS232ModBus_V1.Aux.StartAddr + 6;
       #AteqLeakTest_TCP2RS232ModBus_V1.CTRL_IN_ProgNo := #AteqLeakTest_TCP2RS232ModBus_V1.Aux.StartAddr + 12;
       #AteqLeakTest_TCP2RS232ModBus_V1.Ctrl_IN_ModBusSlaveNO := #AteqLeakTest_TCP2RS232ModBus_V1.Aux.StartAddr + 20;
       #AteqLeakTest_TCP2RS232ModBus_V1.CTRL_Out_ProgNo := #AteqLeakTest_TCP2RS232ModBus_V1.Aux.StartAddr + 32;
       #AteqLeakTest_TCP2RS232ModBus_V1.CTRL_OUT_OKCounter := #AteqLeakTest_TCP2RS232ModBus_V1.Aux.StartAddr + 34;
       #AteqLeakTest_TCP2RS232ModBus_V1.CTRL_OUT_NOKCounter := #AteqLeakTest_TCP2RS232ModBus_V1.Aux.StartAddr + 38;
       #AteqLeakTest_TCP2RS232ModBus_V1.CTRL_OUT_LastCylceTime := #AteqLeakTest_TCP2RS232ModBus_V1.Aux.StartAddr + 42;
       #AteqLeakTest_TCP2RS232ModBus_V1.CTRL_OUT_Pressure := #AteqLeakTest_TCP2RS232ModBus_V1.Aux.StartAddr + 46;
       #AteqLeakTest_TCP2RS232ModBus_V1.CTRL_OUT_LeakRate := #AteqLeakTest_TCP2RS232ModBus_V1.Aux.StartAddr + 50;
       #AteqLeakTest_TCP2RS232ModBus_V1.Status_PromptValue := #AteqLeakTest_TCP2RS232ModBus_V1.Aux.StartAddr + 60;
       #TCPIP_Client_V3.FBCall_StartAddr := #AteqLeakTest_TCP2RS232ModBus_V1.Aux.StartAddr + 174;
       #TCPIP_Client_V3.FBCall_IndexNO := 1;
   END_IF;
   IF #IFM_O2D22X_TCP_V1.FBCall_StartAddr <> #IFM_O2D22X_TCP_V1.Aux.FBCall_StartAddr
       OR #IFM_O2D22X_TCP_V1.FBCall_IndexNO <> #IFM_O2D22X_TCP_V1.Aux.FBCall_IndexNO THEN
       #IFM_O2D22X_TCP_V1.Aux.FBCall_StartAddr := #IFM_O2D22X_TCP_V1.FBCall_StartAddr;
       #IFM_O2D22X_TCP_V1.Aux.FBCall_IndexNO := #IFM_O2D22X_TCP_V1.FBCall_IndexNO;
       #IFM_O2D22X_TCP_V1.Aux.StartAddr := #IFM_O2D22X_TCP_V1.Aux.FBCall_StartAddr +
       (#IFM_O2D22X_TCP_V1.Aux.FBCall_IndexNO - 1) *
       #IFM_O2D22X_TCP_V1.FB_ByteLength;
       #IFM_O2D22X_TCP_V1.TP_Cmd := #IFM_O2D22X_TCP_V1.Aux.StartAddr + 6;
       #IFM_O2D22X_TCP_V1.TP_Status := #IFM_O2D22X_TCP_V1.Aux.StartAddr + 8;
       #IFM_O2D22X_TCP_V1.CTRL_IN_ProgNo := #IFM_O2D22X_TCP_V1.Aux.StartAddr + 14;
       #IFM_O2D22X_TCP_V1.CTRL_IN_DigitOutPutsOKBit := #IFM_O2D22X_TCP_V1.Aux.StartAddr + 16;
       #IFM_O2D22X_TCP_V1.CTRL_Out_ProgNo := #IFM_O2D22X_TCP_V1.Aux.StartAddr + 32;
       #IFM_O2D22X_TCP_V1.CTRL_OUT_OKCounter := #IFM_O2D22X_TCP_V1.Aux.StartAddr + 34;
       #IFM_O2D22X_TCP_V1.CTRL_OUT_NOKCounter := #IFM_O2D22X_TCP_V1.Aux.StartAddr + 38;
       #IFM_O2D22X_TCP_V1.CTRL_OUT_LastCylceTime := #IFM_O2D22X_TCP_V1.Aux.StartAddr + 42;
       #IFM_O2D22X_TCP_V1.CTRL_OUT_DigitOutPutsOKBit := #IFM_O2D22X_TCP_V1.Aux.StartAddr + 46;
       #IFM_O2D22X_TCP_V1.Status_PromptValue := #IFM_O2D22X_TCP_V1.Aux.StartAddr + 50;
       #TCPIP_Client_V3.FBCall_StartAddr := #IFM_O2D22X_TCP_V1.Aux.StartAddr + 110;
       #TCPIP_Client_V3.FBCall_IndexNO := 1;
   END_IF;
   IF #Analog_IN_V4.FBCall_StartAddr <> #Analog_IN_V4.Aux.FBCall_StartAddr
       OR #Analog_IN_V4.FBCall_IndexNO <> #Analog_IN_V4.Aux.FBCall_IndexNO THEN
       #Analog_IN_V4.Aux.FBCall_StartAddr := #Analog_IN_V4.FBCall_StartAddr;
       #Analog_IN_V4.Aux.FBCall_IndexNO := #Analog_IN_V4.FBCall_IndexNO;
       #Analog_IN_V4.Aux.StartAddr := #Analog_IN_V4.Aux.FBCall_StartAddr +
       (#Analog_IN_V4.Aux.FBCall_IndexNO - 1) *
       #Analog_IN_V4.FB_ByteLength;
       #Analog_IN_V4.TP_Cmd := #Analog_IN_V4.Aux.StartAddr + 28;
       #Analog_IN_V4.CTRL_IN_TP_AI_Gain := #Analog_IN_V4.Aux.StartAddr + 34;
       #Analog_IN_V4.CTRL_IN_TP_AI_OffSet := #Analog_IN_V4.Aux.StartAddr + 38;
       #Analog_IN_V4.CTRL_IN_TP_PreSetValue := #Analog_IN_V4.Aux.StartAddr + 42;
       #Analog_IN_V4.CTRL_IN_TP_ActualAI_1 := #Analog_IN_V4.Aux.StartAddr + 46;
       #Analog_IN_V4.CTRL_IN_TP_ActualAI_2 := #Analog_IN_V4.Aux.StartAddr + 50;
       #Analog_IN_V4.CTRL_IN_TP_ActualAI_Value1 := #Analog_IN_V4.Aux.StartAddr + 54;
       #Analog_IN_V4.CTRL_IN_TP_ActualAI_Value2 := #Analog_IN_V4.Aux.StartAddr + 58;
       #Analog_IN_V4.CTRL_OUT_Cur_Val_Out := #Analog_IN_V4.Aux.StartAddr + 80;
       #Analog_IN_V4.CTRL_OUT_TrigerValue := #Analog_IN_V4.Aux.StartAddr + 84;
       #Analog_IN_V4.CTRL_OUT_TrigerValue_Array := #Analog_IN_V4.Aux.StartAddr + 88;
       #Analog_IN_V4.CTRL_OUT_TrigerTPColorStatus_Array := #Analog_IN_V4.Aux.StartAddr + 92;
       #Analog_IN_V4.CTRL_OUT_TrigerCounter := #Analog_IN_V4.Aux.StartAddr + 96;
   END_IF;
END_FUNCTION_BLOCK

FUNCTION_BLOCK "FB5008_CycleTime"   // FB5008, SCL
{ S7_Optimized_Access := 'TRUE' }
// ============================================================
//  Block: FB5008_CycleTime
//  ============================================================
//  编号：FB5008
//  原始语言：LAD（规则翻译为 SCL）
//  含义：由 LAD/FBD 网络折叠生成的等效 SCL，导入前请人工复核
   VAR_INPUT
      StepStart : Bool;   // 输入参数
   END_VAR
   VAR
      CycleTime_Net : Time;   // 静态变量
      CycleTime_Total : Time;   // 静态变量
      Aux : Struct   // 静态变量
         StartPls : Bool;   // 静态变量
         EndPls : Bool;   // 静态变量
         sp : Byte;   // 静态变量
         StartTime : Time_Of_Day;   // 静态变量
         LastEndTime : Time_Of_Day;   // 静态变量
      END_STRUCT;
   END_VAR
   VAR_TEMP
      StepPls : Bool;   // 临时变量
      RetVal : Int;   // 临时变量
   END_VAR
BEGIN

   // ---------- 网络 1 ----------
   // 含义：将 "DB1001_SysMode".Sys_Time.CurPLCTime; (* T_CONV DTL → Time_Of_Day *) 赋给 "SyS_Time"
   "SyS_Time" := DTL_TO_TOD("DB1001_SysMode".Sys_Time.CurPLCTime);

   // ---------- 网络 2 ----------
   // 标题：计算机器运行时间
   // 含义：条件 #StepStart AND NOT (#Aux.StartPls) 成立时，将 "SyS_Time" 传送到 #Aux.StartTime
   IF #StepStart AND NOT (#Aux.StartPls) THEN
       #Aux.StartTime := "SyS_Time";
   END_IF;
   // 含义：当 #StepStart 为 TRUE 时置位 #Aux.StartPls，否则复位（触点→线圈）
   IF #StepStart THEN
       #Aux.StartPls := TRUE;
   ELSE
       #Aux.StartPls := FALSE;
   END_IF;
   // 含义：条件 #StepStart 成立时，将 ("SyS_Time" - #Aux.StartTime) 传送到 #CycleTime_Net
   IF #StepStart THEN
       #CycleTime_Net := ("SyS_Time" - #Aux.StartTime);
   END_IF;

   // ---------- 网络 3 ----------
   // 标题：计算总时间
   // 含义：条件 NOT (#StepStart) AND NOT (#Aux.EndPls) 成立时，将 ("SyS_Time" - #Aux.LastEndTime) 传送到 #CycleTime_Total
   IF NOT (#StepStart) AND NOT (#Aux.EndPls) THEN
       #CycleTime_Total := ("SyS_Time" - #Aux.LastEndTime);
   END_IF;
   // 含义：条件 NOT (#StepStart) AND NOT (#Aux.EndPls) 成立时，将 "SyS_Time" 传送到 #Aux.LastEndTime
   IF NOT (#StepStart) AND NOT (#Aux.EndPls) THEN
       #Aux.LastEndTime := "SyS_Time";
   END_IF;
   // 含义：当 NOT (#StepStart) 为 TRUE 时置位 #Aux.EndPls，否则复位（触点→线圈）
   IF NOT (#StepStart) THEN
       #Aux.EndPls := TRUE;
   ELSE
       #Aux.EndPls := FALSE;
   END_IF;

   // ---------- 网络 4 ----------
   // （空白网络）
END_FUNCTION_BLOCK

ORGANIZATION_BLOCK "OB1Main"   // OB1, LAD, ProgramCycle
TITLE = "Main Program Sweep (Cycle)"
{ S7_Optimized_Access := 'TRUE' }
VERSION : 0.1
BEGIN

REGION Network 1: "DB_StdSignal"
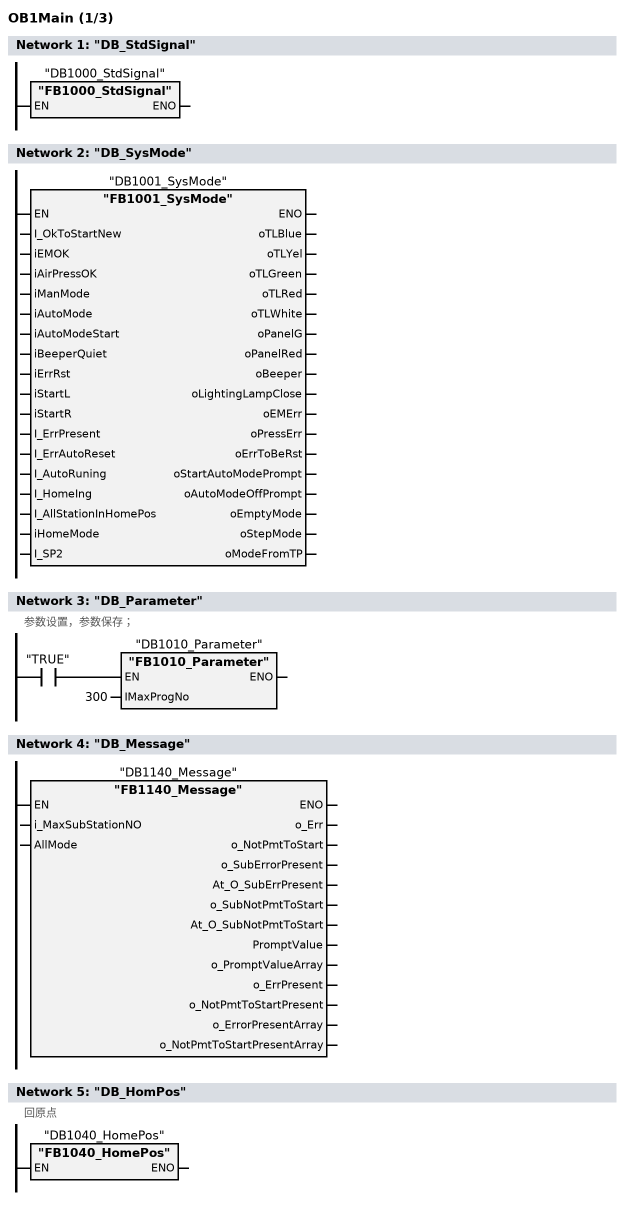
   RUNG wire#powerrail
      "DB1000_StdSignal"()
   END_RUNG
   // the same network as SCL:
   "DB1000_StdSignal"();   // "FB1000_StdSignal"
END_REGION

REGION Network 2: "DB_SysMode"
   RUNG wire#powerrail
      "DB1001_SysMode"(I_OkToStartNew :=, iEMOK :=, iAirPressOK :=, iManMode :=, iAutoMode :=, iAutoModeStart :=, iBeeperQuiet :=, iErrRst :=, iStartL :=, iStartR :=, I_ErrPresent :=, I_ErrAutoReset :=, I_AutoRuning :=, I_HomeIng :=, I_AllStationInHomePos :=, iHomeMode :=, I_SP2 :=, oTLBlue =>, oTLYel =>, oTLGreen =>, oTLRed =>, oTLWhite =>, oPanelG =>, oPanelRed =>, oBeeper =>, oLightingLampClose =>, oEMErr =>, oPressErr =>, oErrToBeRst =>, oStartAutoModePrompt =>, oAutoModeOffPrompt =>, oEmptyMode =>, oStepMode =>, oModeFromTP =>)
   END_RUNG
   // the same network as SCL:
   "DB1001_SysMode"();   // "FB1001_SysMode"
END_REGION

REGION Network 3: "DB_Parameter"
   // 参数设置，参数保存；
   RUNG wire#powerrail
      Contact( "TRUE" )
      "DB1010_Parameter"(IMaxProgNo := 300)
   END_RUNG
   // the same network as SCL:
   IF "TRUE" THEN
       "DB1010_Parameter"(IMaxProgNo := 300);   // "FB1010_Parameter"
   END_IF;
END_REGION

REGION Network 4: "DB_Message"
   RUNG wire#powerrail
      "DB1140_Message"(o_Err =>, o_NotPmtToStart =>, o_SubErrorPresent =>, o_SubNotPmtToStart =>, PromptValue =>, o_PromptValueArray =>, i_MaxSubStationNO :=, AllMode :=, At_O_SubErrPresent =>, At_O_SubNotPmtToStart =>, o_ErrPresent =>, o_NotPmtToStartPresent =>, o_ErrorPresentArray =>, o_NotPmtToStartPresentArray =>)
   END_RUNG
   // the same network as SCL:
   "DB1140_Message"();   // "FB1140_Message"
END_REGION

REGION Network 5: "DB_HomPos"
   // 回原点
   RUNG wire#powerrail
      "DB1040_HomePos"()
   END_RUNG
   // the same network as SCL:
   "DB1040_HomePos"();   // "FB1040_HomePos"
END_REGION

REGION Network 6: "DB_AutoStep"
   // 自动过程
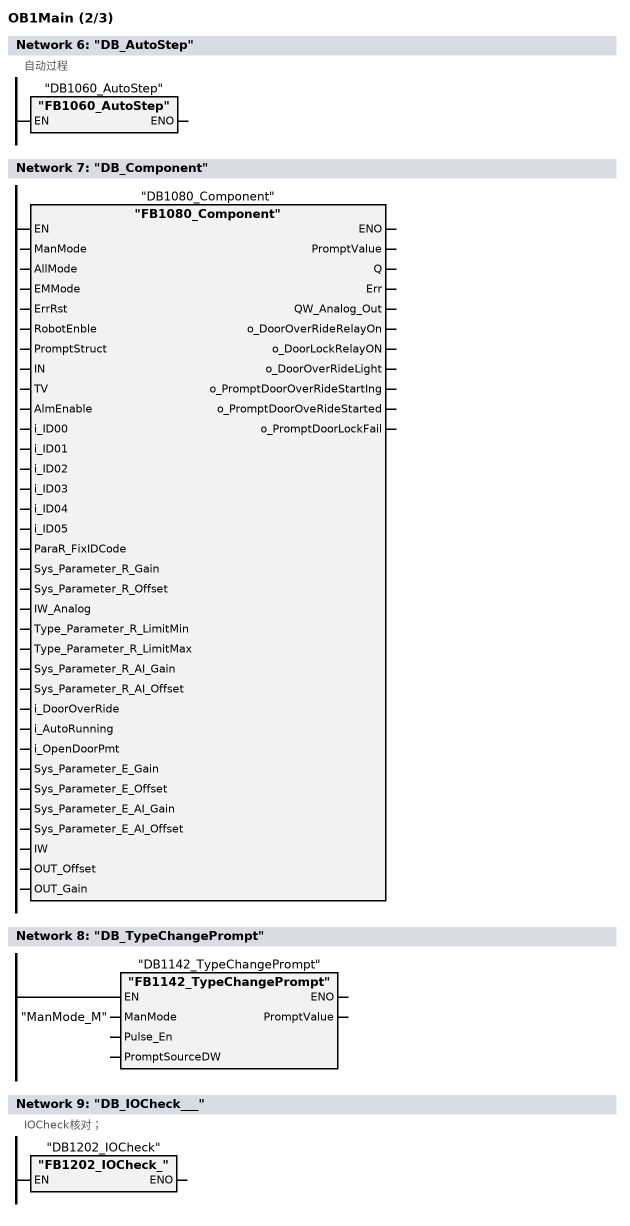
   RUNG wire#powerrail
      "DB1060_AutoStep"()
   END_RUNG
   // the same network as SCL:
   "DB1060_AutoStep"();   // "FB1060_AutoStep"
END_REGION

REGION Network 7: "DB_Component"
   RUNG wire#powerrail
      "DB1080_Component"(ManMode :=, AllMode :=, EMMode :=, ErrRst :=, RobotEnble :=, PromptStruct :=, IN :=, TV :=, AlmEnable :=, i_ID00 :=, i_ID01 :=, i_ID02 :=, i_ID03 :=, i_ID04 :=, i_ID05 :=, ParaR_FixIDCode :=, Sys_Parameter_R_Gain :=, Sys_Parameter_R_Offset :=, IW_Analog :=, Type_Parameter_R_LimitMin :=, Type_Parameter_R_LimitMax :=, Sys_Parameter_R_AI_Gain :=, Sys_Parameter_R_AI_Offset :=, i_DoorOverRide :=, i_AutoRunning :=, i_OpenDoorPmt :=, PromptValue =>, Q =>, Err =>, QW_Analog_Out =>, o_DoorOverRideRelayOn =>, o_DoorLockRelayON =>, o_DoorOverRideLight =>, o_PromptDoorOverRideStartIng =>, o_PromptDoorOveRideStarted =>, o_PromptDoorLockFail =>, Sys_Parameter_E_Gain :=, Sys_Parameter_E_Offset :=, Sys_Parameter_E_AI_Gain :=, Sys_Parameter_E_AI_Offset :=, IW :=, OUT_Offset :=, OUT_Gain :=)
   END_RUNG
   // the same network as SCL:
   "DB1080_Component"();   // "FB1080_Component"
END_REGION

REGION Network 8: "DB_TypeChangePrompt"
   RUNG wire#powerrail
      "DB1142_TypeChangePrompt"(ManMode := "ManMode_M", Pulse_En :=, PromptSourceDW :=, PromptValue =>)
   END_RUNG
   // the same network as SCL:
   "DB1142_TypeChangePrompt"(ManMode := "ManMode_M");   // "FB1142_TypeChangePrompt"
END_REGION

REGION Network 9: "DB_IOCheck___"
   // IOCheck核对；
   RUNG wire#powerrail
      "DB1202_IOCheck"()
   END_RUNG
   // the same network as SCL:
   "DB1202_IOCheck"();   // "FB1202_IOCheck_"
END_REGION

REGION Network 10: "DB_Register"
   // 用于计算HMI界面变量的地址
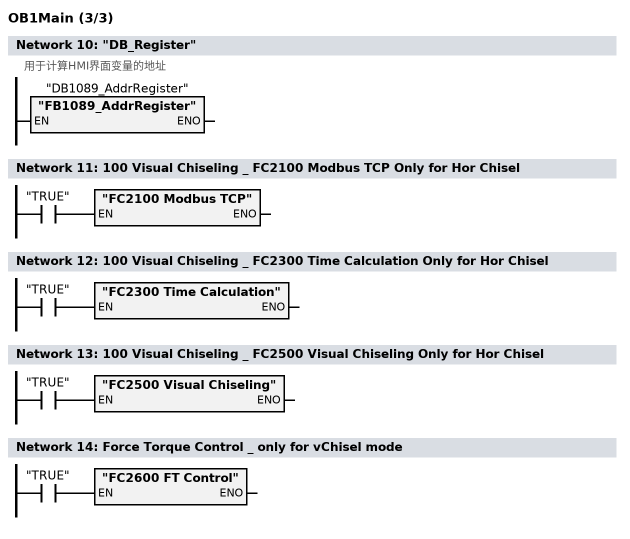
   RUNG wire#powerrail
      "DB1089_AddrRegister"()
   END_RUNG
   // the same network as SCL:
   "DB1089_AddrRegister"();   // "FB1089_AddrRegister"
END_REGION

REGION Network 11: 100 Visual Chiseling _ FC2100 Modbus TCP Only for Hor Chisel
   RUNG wire#powerrail
      Contact( "TRUE" )
      "FC2100 Modbus TCP"()
   END_RUNG
   // the same network as SCL:
   IF "TRUE" THEN "FC2100 Modbus TCP"(); END_IF;
END_REGION

REGION Network 12: 100 Visual Chiseling _ FC2300 Time Calculation Only for Hor Chisel
   RUNG wire#powerrail
      Contact( "TRUE" )
      "FC2300 Time Calculation"()
   END_RUNG
   // the same network as SCL:
   IF "TRUE" THEN "FC2300 Time Calculation"(); END_IF;
END_REGION

REGION Network 13: 100 Visual Chiseling _ FC2500 Visual Chiseling Only for Hor Chisel
   RUNG wire#powerrail
      Contact( "TRUE" )
      "FC2500 Visual Chiseling"()
   END_RUNG
   // the same network as SCL:
   IF "TRUE" THEN "FC2500 Visual Chiseling"(); END_IF;
END_REGION

REGION Network 14: Force Torque Control _ only for vChisel mode
   RUNG wire#powerrail
      Contact( "TRUE" )
      "FC2600 FT Control"()
   END_RUNG
   // the same network as SCL:
   IF "TRUE" THEN "FC2600 FT Control"(); END_IF;
END_REGION
END_ORGANIZATION_BLOCK

ORGANIZATION_BLOCK "OB30_Cyclic interrupt"   // OB30, LAD, CyclicInterrupt
{ S7_Optimized_Access := 'TRUE' }
VERSION : 0.1
   VAR_INPUT
      Initial_Call : Bool;   // Initial call of this OB
      Event_Count : Int;   // Events discarded
   END_VAR
   VAR_TEMP
      PromptForce : Real;
      Temp_ForceNum : Bool;
   END_VAR
   VAR_TEMP   // added for the SCL form of the ladder/FBD networks
      _w1 : Bool;
      _w2 : Bool;
   END_VAR
BEGIN

REGION Network 1: HorDrill Prompt Value Calculation_Not Visual Chiseling Mode
   // GBH2-26 G2  Y=1177.7X-278.46
   // GDB20-160   Y=1560X+36
   // GDB18V Y=1312X+45.4
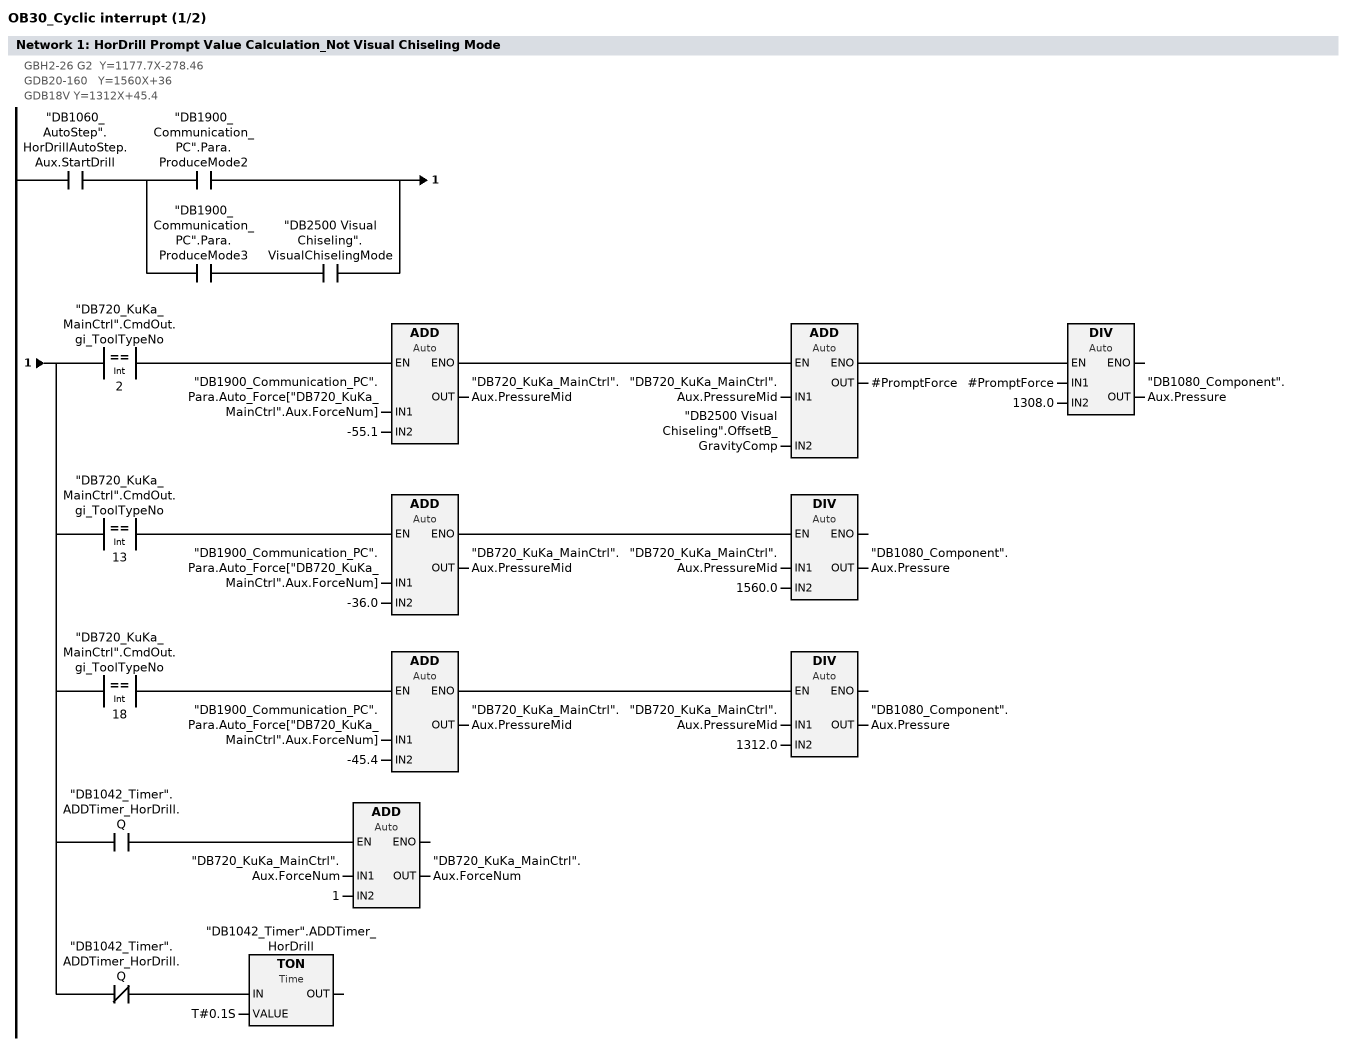
   #_w1 := "DB1060_AutoStep".HorDrillAutoStep.Aux.StartDrill AND ("DB1900_Communication_PC".Para.ProduceMode2 OR ("DB1900_Communication_PC".Para.ProduceMode3 AND "DB2500 Visual Chiseling".VisualChiselingMode));
   IF #_w1 AND ("DB720_KuKa_MainCtrl".CmdOut.gi_ToolTypeNo = 2) THEN
       "DB720_KuKa_MainCtrl".Aux.PressureMid := "DB1900_Communication_PC".Para.Auto_Force["DB720_KuKa_MainCtrl".Aux.ForceNum] + (-55.1);
       #PromptForce := "DB720_KuKa_MainCtrl".Aux.PressureMid + "DB2500 Visual Chiseling".OffsetB_GravityComp;
       "DB1080_Component".Aux.Pressure := #PromptForce / 1308.0;
   END_IF;
   IF #_w1 AND ("DB720_KuKa_MainCtrl".CmdOut.gi_ToolTypeNo = 13) THEN
       "DB720_KuKa_MainCtrl".Aux.PressureMid := "DB1900_Communication_PC".Para.Auto_Force["DB720_KuKa_MainCtrl".Aux.ForceNum] + (-36.0);
       "DB1080_Component".Aux.Pressure := "DB720_KuKa_MainCtrl".Aux.PressureMid / 1560.0;
   END_IF;
   IF #_w1 AND ("DB720_KuKa_MainCtrl".CmdOut.gi_ToolTypeNo = 18) THEN
       "DB720_KuKa_MainCtrl".Aux.PressureMid := "DB1900_Communication_PC".Para.Auto_Force["DB720_KuKa_MainCtrl".Aux.ForceNum] + (-45.4);
       "DB1080_Component".Aux.Pressure := "DB720_KuKa_MainCtrl".Aux.PressureMid / 1312.0;
   END_IF;
   IF #_w1 AND "DB1042_Timer".ADDTimer_HorDrill.Q THEN
       "DB720_KuKa_MainCtrl".Aux.ForceNum := "DB720_KuKa_MainCtrl".Aux.ForceNum + 1;
   END_IF;
   "DB1042_Timer".ADDTimer_HorDrill.TON(IN := #_w1 AND NOT "DB1042_Timer".ADDTimer_HorDrill.Q, PT := T#0.1S);   // TON coil
END_REGION

REGION Network 2: DownDrill Prompt Value Calculation
   // GBH2-26 G2  Y=1177.7X-278.46
   // GDB20-160   Y=1274.3X-51.929
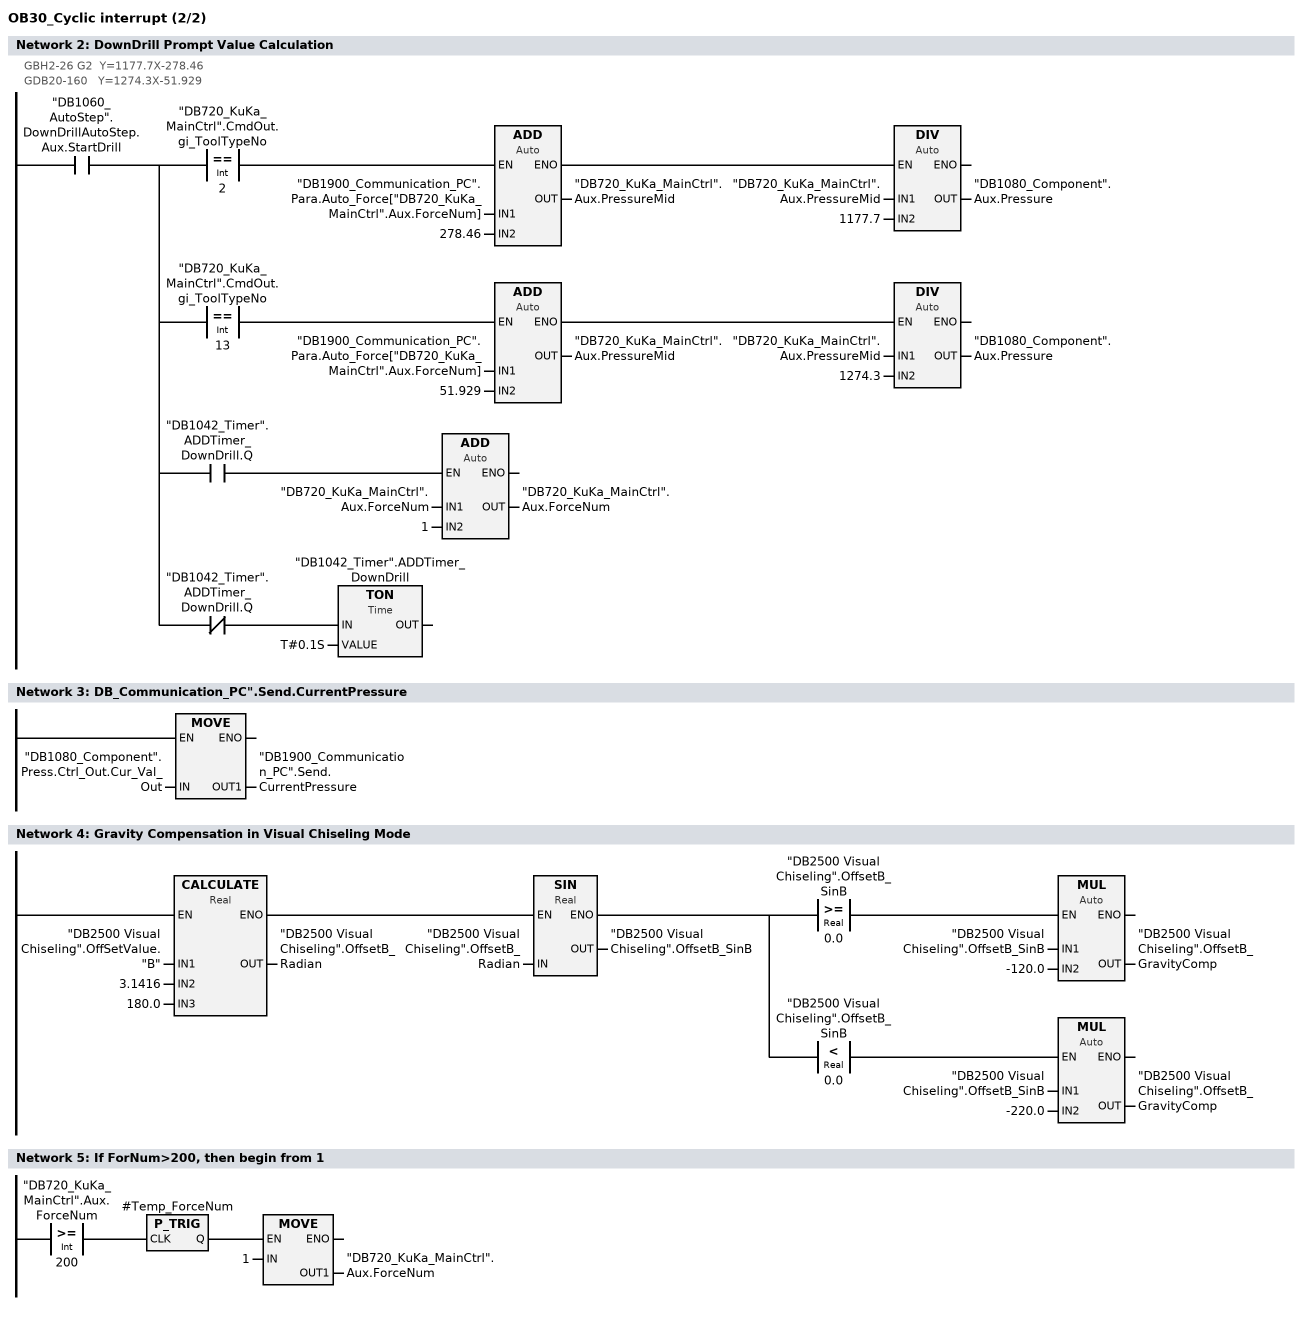
   IF "DB1060_AutoStep".DownDrillAutoStep.Aux.StartDrill AND ("DB720_KuKa_MainCtrl".CmdOut.gi_ToolTypeNo = 2) THEN
       "DB720_KuKa_MainCtrl".Aux.PressureMid := "DB1900_Communication_PC".Para.Auto_Force["DB720_KuKa_MainCtrl".Aux.ForceNum] + 278.46;
       "DB1080_Component".Aux.Pressure := "DB720_KuKa_MainCtrl".Aux.PressureMid / 1177.7;
   END_IF;
   IF "DB1060_AutoStep".DownDrillAutoStep.Aux.StartDrill AND ("DB720_KuKa_MainCtrl".CmdOut.gi_ToolTypeNo = 13) THEN
       "DB720_KuKa_MainCtrl".Aux.PressureMid := "DB1900_Communication_PC".Para.Auto_Force["DB720_KuKa_MainCtrl".Aux.ForceNum] + 51.929;
       "DB1080_Component".Aux.Pressure := "DB720_KuKa_MainCtrl".Aux.PressureMid / 1274.3;
   END_IF;
   IF "DB1060_AutoStep".DownDrillAutoStep.Aux.StartDrill AND "DB1042_Timer".ADDTimer_DownDrill.Q THEN
       "DB720_KuKa_MainCtrl".Aux.ForceNum := "DB720_KuKa_MainCtrl".Aux.ForceNum + 1;
   END_IF;
   "DB1042_Timer".ADDTimer_DownDrill.TON(IN := "DB1060_AutoStep".DownDrillAutoStep.Aux.StartDrill AND NOT "DB1042_Timer".ADDTimer_DownDrill.Q, PT := T#0.1S);   // TON coil
END_REGION

REGION Network 3: DB_Communication_PC".Send.CurrentPressure
   RUNG wire#powerrail
      Move(in := "DB1080_Component".Press.Ctrl_Out.Cur_Val_Out, out1 => "DB1900_Communication_PC".Send.CurrentPressure)
   END_RUNG
   // the same network as SCL:
   "DB1900_Communication_PC".Send.CurrentPressure := "DB1080_Component".Press.Ctrl_Out.Cur_Val_Out;
END_REGION

REGION Network 4: Gravity Compensation in Visual Chiseling Mode
   "DB2500 Visual Chiseling".OffsetB_Radian := ("DB2500 Visual Chiseling".OffSetValue."B"*3.1416)/180.0;
   "DB2500 Visual Chiseling".OffsetB_SinB := SIN("DB2500 Visual Chiseling".OffsetB_Radian);
   IF "DB2500 Visual Chiseling".OffsetB_SinB >= 0.0 THEN
       "DB2500 Visual Chiseling".OffsetB_GravityComp := "DB2500 Visual Chiseling".OffsetB_SinB * (-120.0);
   END_IF;
   IF "DB2500 Visual Chiseling".OffsetB_SinB < 0.0 THEN
       "DB2500 Visual Chiseling".OffsetB_GravityComp := "DB2500 Visual Chiseling".OffsetB_SinB * (-220.0);
   END_IF;
END_REGION

REGION Network 5: If ForNum>200, then begin from 1
   RUNG wire#powerrail
      { S7_Templates := "SrcType := Int" } GE_Contact(in1 := "DB720_KuKa_MainCtrl".Aux.ForceNum, in2 := 200)
      P_Trig( #Temp_ForceNum )
      Move(in := 1, out1 => "DB720_KuKa_MainCtrl".Aux.ForceNum)
   END_RUNG
   // the same network as SCL:
   #_w1 := "DB720_KuKa_MainCtrl".Aux.ForceNum >= 200;
   #_w2 := #_w1 AND NOT #Temp_ForceNum;   // rising edge
   #Temp_ForceNum := #_w1;
   IF #_w2 THEN "DB720_KuKa_MainCtrl".Aux.ForceNum := 1; END_IF;
END_REGION
END_ORGANIZATION_BLOCK

// folder: 001_KL_Standard_FB

FUNCTION_BLOCK "FB950_SDTimer"   // FB950, SCL
{ S7_Optimized_Access := 'TRUE' }
// ============================================================
//  Block: FB950_SDTimer
//  ============================================================
//  编号：FB950
//  原始语言：LAD（规则翻译为 SCL）
//  含义：由 LAD/FBD 网络折叠生成的等效 SCL，导入前请人工复核
   VAR_INPUT
      TV : Time;   // 设置时间(1ms)
   END_VAR
   VAR_IN_OUT
      IN : Bool;   // 输入输出参数
      Q : Bool;   // 输入输出参数
   END_VAR
   VAR
      TempSystime : Time;   // 静态变量
      AtTempDint1 : Time_Of_Day;   // 静态变量
   END_VAR
BEGIN
END_FUNCTION_BLOCK

FUNCTION_BLOCK "FB951_SDTimerV2"   // FB951, SCL
{ S7_Optimized_Access := 'TRUE' }
// ============================================================
//  Block: FB951_SDTimerV2
//  ============================================================
//  编号：FB951
//  原始语言：LAD（规则翻译为 SCL）
//  含义：由 LAD/FBD 网络折叠生成的等效 SCL，导入前请人工复核
   VAR_INPUT
      IN : Bool;   // 开始定时
      TV : Time;   // 设置时间(1ms)
   END_VAR
   VAR_OUTPUT
      Q : Bool;   // 时间到达
   END_VAR
   VAR
      StartTime : Time;   // 开始时间
      AtStartTime : Time_Of_Day;   // 静态变量
      ET : Time;   // 过去的时间
      IN_EDGE : Bool;   // 边沿记忆
   END_VAR
BEGIN
END_FUNCTION_BLOCK

FUNCTION_BLOCK "FB1000_StdSignal"   // FB1000, SCL
{ S7_Optimized_Access := 'TRUE' }
// ============================================================
//  Block: FB1000_StdSignal
//  ============================================================
//  编号：FB1000
//  原始语言：LAD（规则翻译为 SCL）
//  含义：由 LAD/FBD 网络折叠生成的等效 SCL，导入前请人工复核
   VAR
      PLS : Struct   // 静态变量
         PS02 : Bool;   // 静态变量
         PS05 : Bool;   // 静态变量
         PS10 : Bool;   // 静态变量
         PS01 : Bool;   // 静态变量
         PromptRenewPls : Bool;   // 静态变量
         InitialPls : Bool;   // 静态变量
      END_STRUCT;
      RectWave : Struct   // 静态变量
         Wave02 : Bool;   // 200ms ON,200ms OFF.
         Wave05 : Bool;   // 500ms ON,500ms OFF.
         Wave10 : Bool;   // 1s ON,1s OFF.
         Beeper : Bool;   // 静态变量
      END_STRUCT;
      PowerOn : Bool;   // 静态变量
      LampTest : Bool;   // 静态变量
      AlwaysOn : Bool;   // 静态变量
      TimerStruct : Struct   // 静态变量
         T100ms脉冲定时 : IEC_TIMER;   // 静态变量
         T200ms脉冲定时 : IEC_TIMER;   // 静态变量
         T500ms脉冲定时 : IEC_TIMER;   // 静态变量
         T1s脉冲定时 : IEC_TIMER;   // 静态变量
         PromptRenewPls : IEC_TIMER;   // 静态变量
         T200ms方波定时1 : IEC_TIMER;   // 静态变量
         T200ms方波定时2 : IEC_TIMER;   // 静态变量
         T500ms方波定时1 : IEC_TIMER;   // 静态变量
         T500ms方波定时2 : IEC_TIMER;   // 静态变量
         T1S方波定时1 : IEC_TIMER;   // 静态变量
         T1S方波定时2 : IEC_TIMER;   // 静态变量
         T_PowerOn1 : IEC_TIMER;   // 静态变量
         T_PowerOn2 : IEC_TIMER;   // 静态变量
         Beeper1 : IEC_TIMER;   // 静态变量
         Beeper2 : IEC_TIMER;   // 静态变量
      END_STRUCT;
      PT : Time;   // 静态变量
      ET : Time;   // 静态变量
      IN : Bool;   // 静态变量
      Q : Bool;   // 静态变量
   END_VAR
BEGIN
END_FUNCTION_BLOCK

FUNCTION_BLOCK "FB1021_Prompt_Object"   // FB1021, SCL
{ S7_Optimized_Access := 'TRUE' }
// ============================================================
//  Block: FB1021_Prompt_Object
//  ============================================================
//  编号：FB1021
//  原始语言：SCL（规则翻译为 SCL）
//  含义：由 LAD/FBD 网络折叠生成的等效 SCL，导入前请人工复核
   VAR_INPUT
      Pulse_En : Bool;   // 更新脉冲
      PromptSourceDW : DWord;   // 输入参数
   END_VAR
   VAR_OUTPUT
      PromptValue : Int;   // 用于触摸屏
   END_VAR
   VAR
      CycleTime : Int;   // 循环次数计数
      PromptValueBake : Int;   // 提示值暂存；
      ShiftBake : Int;   // 静态变量
   END_VAR
BEGIN
END_FUNCTION_BLOCK

FUNCTION_BLOCK "FB1022_Prompt_ObjectV2"   // FB1022, SCL
{ S7_Optimized_Access := 'TRUE' }
// ============================================================
//  Block: FB1022_Prompt_ObjectV2
//  ============================================================
//  编号：FB1022
//  原始语言：SCL（规则翻译为 SCL）
//  含义：由 LAD/FBD 网络折叠生成的等效 SCL，导入前请人工复核
   VAR_INPUT
      PromptStruct : Struct   // 输入参数
         Info : Struct   // 输入参数
            bit0 : Bool;   // 输入参数
            bit1 : Bool;   // 输入参数
            bit2 : Bool;   // 输入参数
            bit3 : Bool;   // 输入参数
            bit4 : Bool;   // 输入参数
            bit5 : Bool;   // 输入参数
            bit6 : Bool;   // 输入参数
            bit7 : Bool;   // 输入参数
            bit8 : Bool;   // 输入参数
            bit9 : Bool;   // 输入参数
            bit10 : Bool;   // 输入参数
            bit11 : Bool;   // 输入参数
            bit12 : Bool;   // 输入参数
            bit13 : Bool;   // 输入参数
            bit14 : Bool;   // 输入参数
            bit15 : Bool;   // 输入参数
            bit16 : Bool;   // 输入参数
            bit17 : Bool;   // 输入参数
            bit18 : Bool;   // 输入参数
            bit19 : Bool;   // 输入参数
            bit20 : Bool;   // 输入参数
            bit21 : Bool;   // 输入参数
            bit22 : Bool;   // 输入参数
            bit23 : Bool;   // 输入参数
            bit24 : Bool;   // 输入参数
            bit25 : Bool;   // 输入参数
            bit26 : Bool;   // 输入参数
            bit27 : Bool;   // 输入参数
            bit28 : Bool;   // 输入参数
            bit29 : Bool;   // 输入参数
            bit30 : Bool;   // 输入参数
            bit31 : Bool;   // 输入参数
         END_STRUCT;
         Err : Struct   // 输入参数
            bit0 : Bool;   // 输入参数
            bit1 : Bool;   // 输入参数
            bit2 : Bool;   // 输入参数
            bit3 : Bool;   // 输入参数
            bit4 : Bool;   // 输入参数
            bit5 : Bool;   // 输入参数
            bit6 : Bool;   // 输入参数
            bit7 : Bool;   // 输入参数
            bit8 : Bool;   // 输入参数
            bit9 : Bool;   // 输入参数
            bit10 : Bool;   // 输入参数
            bit11 : Bool;   // 输入参数
            bit12 : Bool;   // 输入参数
            bit13 : Bool;   // 输入参数
            bit14 : Bool;   // 输入参数
            bit15 : Bool;   // 输入参数
            bit16 : Bool;   // 输入参数
            bit17 : Bool;   // 输入参数
            bit18 : Bool;   // 输入参数
            bit19 : Bool;   // 输入参数
            bit20 : Bool;   // 输入参数
            bit21 : Bool;   // 输入参数
            bit22 : Bool;   // 输入参数
            bit23 : Bool;   // 输入参数
            bit24 : Bool;   // 输入参数
            bit25 : Bool;   // 输入参数
            bit26 : Bool;   // 输入参数
            bit27 : Bool;   // 输入参数
            bit28 : Bool;   // 输入参数
            bit29 : Bool;   // 输入参数
            bit30 : Bool;   // 输入参数
            bit31 : Bool;   // 输入参数
         END_STRUCT;
      END_STRUCT;
      AtPromptStruct : Struct   // 输入参数
         Info : DWord;   // 输入参数
         Err : DWord;   // 输入参数
      END_STRUCT;
   END_VAR
   VAR_OUTPUT
      PromptValue : Int;   // 用于触摸屏
   END_VAR
   VAR
      CycleTime : Int;   // 循环次数计数
      PromptValueBake : Int;   // 提示值暂存；
      ShiftBake : Int;   // 静态变量
   END_VAR
BEGIN
END_FUNCTION_BLOCK

FUNCTION_BLOCK "FB1141_Prompt"   // FB1141, SCL
{ S7_Optimized_Access := 'TRUE' }
// ============================================================
//  Block: FB1141_Prompt
//  ============================================================
//  编号：FB1141
//  原始语言：SCL（规则翻译为 SCL）
//  含义：由 LAD/FBD 网络折叠生成的等效 SCL，导入前请人工复核
   VAR_INPUT
      i_MaxSubStationNO : Int := 1;   // 输入参数
      AllMode : Bool;   // 输入参数
   END_VAR
   VAR_OUTPUT
      o_ErrPresent : Bool;   // DB_Err任意一位=On
      o_NotPmtToStartPresent : Bool;   // DB_PromptStartNotPmt及DB_Err任意一位=On
      o_ErrorPresentArray : Array[0..31] of Bool;   // 各子工位存在故障，用于识别各个子站是否需要回原点
      At_o_ErrPresentArray : DWord;   // 输出参数
      o_NotPmtToStartPresentArray : Array[0..31] of Bool;   // 各子工位存在故障，用于识别各个子站是否需要回原点
      At_o_NotPmtToStartPresentArray : DWord;   // 输出参数
      PromptValue : Int;   // 总的提示信息
      o_PromptValueArray : Array[0..31] of Int;   // 各个子工位的提示信息
   END_VAR
   VAR
      Para : Struct   // 静态变量
         StartDBNO : Int := 1146;   // 本程序处理的DB编号起始地址
         DBLoopCounter : Int := 2;   // 0..2,即默认是DB1146~~1148
         DBMessage_Gap : Int := 1000;   // 不同DB消息之间的间隔，当DB区域大于125Byte时，需要加大该值
      END_STRUCT;
      Para_ReserveLength : Struct   // 参数信息，请直接在FB内赋默认值
         DB_PromptFree : Array[0..31] of Int;   // DB1146各个Struct所含的字节长度, 必须是4的整数倍
         DB_PromptStartNotPmt : Array[0..31] of Int;   // DB1147各个Struct所含的字节长度, 必须是4的整数倍
         DB_PromptErr : Array[0..31] of Int;   // DB1148各个Struct所含的字节长度, 必须是4的整数倍
      END_STRUCT;
      At_ParaReserveLength : Array[0..2, 0..31] of Int;   // 内部变量，请勿赋值
      xAux : Struct   // 内部变量，请勿赋值
         AnyBitOnPresentArray : Array[0..2, 0..31] of Bool;   // 静态变量
         AnyBitOnPresent : Array[0..2] of Bool;   // 所有DB中，任意一个DB有一位处于On状态
         o_PromptValueArray : Array[0..2, 0..31] of Int;   // 提示信息
         BakeArray : Array[0..2, 0..31] of Struct   // 内部程序使用,外部不允许操作
            ScanFinished : Bool;   // 扫描完成
            PromptValueBake : Int;   // 静态变量
         END_STRUCT;
         DB_StationShift : Array[0..2] of Int;   // 静态变量
         ParaSubStationStartByteNO : Array[0..2, 0..31] of Int;   // 静态变量
         o_W_ErrPresentArray : DWord;   // 值同Output: o_ErrorPresentArray数组
         o_W_NotPmtToStartPresentArray : DWord;   // 静态变量
         DBNO : Int;   // 静态变量
         SubStep : Int;   // 静态变量
         JumpStepNO : Int;   // 静态变量
         SubStation : Int;   // 静态变量
         DBNumber : Int;   // 静态变量
      END_STRUCT;
      At_xAux : Struct   // 静态变量
         AnyBitOnPresentArray : Array[0..2] of DWord;   // 静态变量
      END_STRUCT;
      sp : Array[0..113] of Byte;   // 静态变量
      LastAddr : Int := 1198;   // 静态变量
   END_VAR
BEGIN
END_FUNCTION_BLOCK

FUNCTION_BLOCK "FB1200_std_Switch"   // FB1200, SCL
{ S7_Optimized_Access := 'TRUE' }
// ============================================================
//  Block: FB1200_std_Switch
//  ============================================================
//  编号：FB1200
//  原始语言：LAD（规则翻译为 SCL）
//  含义：由 LAD/FBD 网络折叠生成的等效 SCL，导入前请人工复核
   VAR_IN_OUT
      CylinderCmd : Struct   // 输入输出参数
         ExtTPPB : Bool;   // 气缸名1
         RetTPPB : Bool;   // 气缸名1
         ExtPmt : Bool;   // 气缸名1
         RetPmt : Bool;   // 气缸名1
         IExtPos : Bool;   // 气缸名1
         IRetPos : Bool;   // 气缸名1
         TPSP1 : Bool;   // 气缸名1
         VentValveTPPB : Bool;   // 气缸名1
         ExtEVT : Bool;   // 气缸名1
         RetEVT : Bool;   // 气缸名1
         ExtPos : Bool;   // 气缸名1
         RetPos : Bool;   // 气缸名1
         ExtIng : Bool;   // 气缸名1
         RetIng : Bool;   // 气缸名1
         ExtErr : Bool;   // 气缸名1
         RetErr : Bool;   // 气缸名1
         ExtAuto : Bool;   // 气缸名1
         RetAuto : Bool;   // 气缸名1
         VentValveAuto : Bool;   // 气缸名1
         VentValve : Bool;   // 气缸名1
         Moving : Bool;   // 气缸名1
         RegTimer : Int;   // 气缸名1
      END_STRUCT;
   END_VAR
   VAR
      ManMode : Bool;   // 手动模式
      AllMode : Bool;   // 所有模式
      EMMode : Bool;   // 紧急停止模式
      OprNotPmt : Bool;   // 操作被禁止
      ResetAllCmd : Bool;   // 复位所有的动作命令
   END_VAR
BEGIN
END_FUNCTION_BLOCK

FUNCTION_BLOCK "FB1202_IOCheck_"   // FB1202, SCL
{ S7_Optimized_Access := 'TRUE' }
// ============================================================
//  Block: FB1202_IOCheck_
//  ============================================================
//  编号：FB1202
//  原始语言：LAD（规则翻译为 SCL）
//  含义：由 LAD/FBD 网络折叠生成的等效 SCL，导入前请人工复核
   VAR
      Status : Struct   // 静态变量
         Sp0 : Bool;   // 上页
         Sp1 : Bool;   // 下页
         Sp2 : Bool;   // 上页
         Sp3 : Bool;   // 下页
         Sp4 : Bool;   // 静态变量
         Sp5 : Bool;   // 静态变量
         Sp6 : Bool;   // 静态变量
         Sp7 : Bool;   // 静态变量
         InPrePageEnd : Bool;   // In上页到头
         InNextPageEnd : Bool;   // In下页到头
         OutPrePageEnd : Bool;   // Out上页到头
         OutNextPageEnd : Bool;   // Out下页到头
      END_STRUCT;
      AtStatus : Word;   // 静态变量
      TP_Status : Word;   // 静态变量
      In_ByteNo : Int;   // Out当前要显示的Byte编号IB0，ByteNo=0
      Out_ByteNo : Int;   // Out当前要显示的Byte编号IB0，ByteNo=0
      In_ByteNo_X10 : Array[0..7] of Int;   // 用于更新当前显示Input的内容；
      Out_ByteNo_X10 : Array[0..7] of Int;   // 用于更新当前显示OutPut的内容；
      InputMaxByteNo : Int;   // 输入IO最大Byte地址
      InputMinByteNo : Int;   // 输入IO最小Byte地址
      OutputMaxByteNo : Int;   // 输出IO最大Byte地址
      OutputMinByteNo : Int;   // 输出IO最小Byte地址
      Aux : Struct   // 静态变量
         In_IndexNo_Bake : Int;   // Out当前要显示的Byte编号IB0，ByteNo=0
         Out_IndexNo_Bake : Int;   // Out当前要显示的Byte编号IB0，ByteNo=0
      END_STRUCT;
   END_VAR
BEGIN
END_FUNCTION_BLOCK

FUNCTION_BLOCK "FB1210_DPRD_DPWR"   // FB1210, SCL
{ S7_Optimized_Access := 'TRUE' }
// ============================================================
//  Block: FB1210_DPRD_DPWR
//  ============================================================
//  编号：FB1210
//  原始语言：SCL（规则翻译为 SCL）
//  含义：由 LAD/FBD 网络折叠生成的等效 SCL，导入前请人工复核
   VAR_INPUT
      bReadOrWrite : Bool;   // False: To Read Input, True: To Write Output
      IO_Addr : DInt;   // 输入参数
      IO_LenOfByte : DInt;   // 输入参数
   END_VAR
   VAR
      ByteArray : Array[0..255] of Byte;   // 静态变量
      dbNumber_self : Int := 1210;   // 静态变量
   END_VAR
BEGIN
END_FUNCTION_BLOCK

